// TIA Portal project "HR001_PLC_20260509" (V19)

(* hardware
DEVICE "S7-1200 station_1"  SIMATIC 1200-Station
   slot 0: "S7-1200 rack"  Rack  V1.0
   slot 1: "CPU_1200"  CPU 1215C DC/DC/DC  6ES7 215-1AG40-0XB0  V4.4
   slot 2: "DI 16/DQ 16x24VDC_1"  6ES7 223-1BL32-0XB0  V2.0
   slot 3: "DI 16/DQ 16x24VDC_2"  6ES7 223-1BL32-0XB0  V2.0
   slot 4: "DI 16x24VDC_1"  6ES7 221-1BH32-0XB0  V2.0
DEVICE "GSD device_11"  GSD.Device.PN
   slot 0: "机架"  Rack  V1.0
   slot 0: "AG1521Kuka_Big"  KRC4-ProfiNet_3.2  V3.2
      slot 0: "KRC4-ProfiNet_3.2"  KRC4-ProfiNet_3.2
      slot 1: "Interface1"  Interface1
         slot 1: "Port1"  Port1
   slot 2: "512 digital in- and outputs_1"  512 digital in- and outputs  KUKA KR C4 Device IO512
      slot 0: "512 digital in- and outputs"  512 digital in- and outputs
DEVICE "TP"  SIMATIC PC station
   slot 0: "HMI"  Rail  SIMATIC PC-Station  V1.0
      slot 125: "Stationmanager"  Station_Manager  V6.0.4
   slot 1: "HMI_RT_1"  WinCC RT Advanced  6AV2 104-0xxxx-xxxx  16.0.0.0
      slot 33792: "Computer interface"  Host interface
   slot 4: "IE general_1"  IE General  IE_CP  V8.2.0
*)

// ===== PLC "CPU_1200"  CPU 1215C DC/DC/DC =====
// protected blocks, not shown: "FB1003_CR", "FC1003_CR"

VAR_GLOBAL   // PLC tag table "M变量"
   "ManMode_M" AT %M26.0 : Bool;   // 手动模式
   "MastMode_M" AT %M26.1 : Bool;   // 校验模式
   "StepMode_M" AT %M26.2 : Bool;   // 单步模式
   "AutoMode_M" AT %M26.3 : Bool;   // 自动模式
   "EMMode_M" AT %M26.4 : Bool;   // 急停
   "StepPls_M" AT %M26.5 : Bool;   // 单步
   "AutoModeStarted_M" AT %M26.7 : Bool;   // 自动开始
   "ASMode_M" AT %M27.0 : Bool;   // 自动、单步
   "ASMMode_M" AT %M27.1 : Bool;   // 自动、单步、校验模式
   "AllMode_M" AT %M27.2 : Bool;   // 所有模式
   "ErrRst_M" AT %M27.3 : Bool;   // 故障复位
   "ErrRst_M_Auto" AT %M27.4 : Bool;   // 故障复位(系统参数可以设置为自动复位信号)
   "TRUE" AT %M29.0 : Bool;
   "False" AT %M29.1 : Bool;
   "MESConnect" AT %M29.3 : Bool;   // 0单机1联机
   "Debug_True" AT %M29.4 : Bool;   // 调试的时候，临时关闭
   "SyS_Time" AT %MD30 : Time_Of_Day;
   "Tag_1" AT %MW120 : Word;
   "Tag_2" AT %MW108 : Word;
   "Tag_3" AT %MW112 : UInt;
   "Tag_4" AT %M29.5 : Bool;
END_VAR

VAR_GLOBAL   // PLC tag table "PLC_IO"
   "IDoor3Unlocked" AT %I2.0 : Bool;   // 垂直击打门锁未锁定
   "IDoor3Insert" AT %I2.1 : Bool;   // 垂直击打门锁已插入
   "AStation_ToolOn2" AT %I2.5 : Bool;   // A工位夹具 有无检测2
   "AStation_ToolOn1" AT %I2.4 : Bool;   // A工位夹具 有无检测1
   "AStation_IZ03ExtPos" AT %I3.0 : Bool;   // A工位 旋转压紧缸伸出磁开
   "AStation_IZ03RetPos" AT %I3.1 : Bool;   // A工位 旋转压紧缸缩回磁开
   "BStation_ToolOn2" AT %I2.3 : Bool;   // B工位夹具有无检测2
   "BStation_ToolOn1" AT %I2.2 : Bool;   // B工位夹具 有无检测1
   "ICurtainErrRst" AT %I1.0 : Bool;   // 光幕复位按钮
   "IDoorOverRide" AT %I1.1 : Bool;   // 安全门旁路
   "IDoor1Unlocked" AT %I1.2 : Bool;   // 产品上料门锁未锁定
   "IDoor1Insert" AT %I1.3 : Bool;   // 产品上料门锁已插入
   "IDoor2Unlocked" AT %I1.4 : Bool;   // 水平击打门锁未锁定
   "IDoor2Insert" AT %I1.5 : Bool;   // 水平击打门锁已插入
   "IFixtureCode02" AT %I4.0 : Bool;   // 夹具电源快插编码2
   "IFixtureCode03" AT %I4.1 : Bool;   // 夹具电源快插编码3
   "IFixtureIOCode01" AT %I4.2 : Bool;   // 夹具IO快插编码1
   "IFixtureIOCode02" AT %I4.3 : Bool;   // 夹具IO快插编码2
   "IFixtureIOCode03" AT %I4.4 : Bool;   // 夹具IO快插编码3
   "IEMClamp" AT %I4.5 : Bool;   // 夹具侧急停按钮
   "IFixtureStuckSensor" AT %I4.6 : Bool;   // 夹具防卡信号
   "ISp4_7" AT %I4.7 : Bool;
   "IRobotEMOK" AT %I5.1 : Bool;   // 机器人急停按钮OK
   "ICurtainsOK" AT %I0.6 : Bool;   // 光幕OK信号
   "BStation_IZ04RetPos" AT %I2.6 : Bool;   // B工位 旋转压紧缸缩回磁开
   "IZ02RetPos" AT %I3.3 : Bool;   // 辅助气缸缩回磁开
   "IZ07ExtPos" AT %I3.5 : Bool;   // 机器人快换盘夹紧
   "IZ07RetPos" AT %I3.4 : Bool;   // 机器人快换盘松开
   "IToolAtPos" AT %I3.6 : Bool;   // 机器人快换盘在位
   "IFixtureCode01" AT %I3.7 : Bool;   // 夹具电源快插编码1
   "IEMOK" AT %I0.0 : Bool;   // 紧急停止OK
   "IAirPressOK" AT %I0.1 : Bool;   // 总气压检测OK
   "IMan" AT %I0.2 : Bool;   // 手动模式
   "IAuto" AT %I0.3 : Bool;   // 自动模式
   "IAutoModeStart" AT %I0.4 : Bool;   // 自动启动按钮
   "IErrRst" AT %I0.5 : Bool;   // 故障复位按钮
   "BStation_IZ04ExtPos" AT %I2.7 : Bool;   // B工位 旋转压紧缸伸出磁开
   "IZ02ExtPos" AT %I3.2 : Bool;   // 辅助气缸伸出磁开
   "IAllDoorClose" AT %I5.0 : Bool;   // 上电&所有 安全门关闭
   "IEMOK1" AT %I0.7 : Bool;   // 操作盒急停OK
   "ITempErr" AT %I5.2 : Bool;   // 温控器报警
   "IInsideEMOK" AT %I5.3 : Bool;   // 围栏内侧急停信号
   "IInsideEMOK1" AT %I5.4 : Bool;   // 水泥块击打框架急停信号
   "ISp055" AT %I5.5 : Bool;   // 备用
   "ISp056" AT %I5.6 : Bool;   // 备用
   "ISp057" AT %I5.7 : Bool;   // 备用
   "QBeeper" AT %Q0.2 : Bool;   // 蜂鸣器
   "QPanelG" AT %Q0.0 : Bool;   // 绿色运行指示灯
   "QPanelRed" AT %Q0.1 : Bool;   // 故障复位红灯
   "QTLR" AT %Q0.3 : Bool;   // 五色塔灯(红)
   "QTLY" AT %Q0.4 : Bool;   // 五色塔灯(黄)
   "QTLG" AT %Q0.5 : Bool;   // 五色塔灯(绿)
   "QTLB" AT %Q0.6 : Bool;   // 五色塔灯(蓝)
   "QTLW" AT %Q0.7 : Bool;   // 五色塔灯(白)
   "QSpairMode" AT %Q1.0 : Bool;   // 安全门旁路
   "QLampCtr" AT %Q1.1 : Bool;   // 日光灯控制中继（预留）
   "OOpenCamCover" AT %Q1.2 : Bool;   // 打开相机防护罩
   "OCloseCamCover" AT %Q1.3 : Bool;   // 关闭相机防护罩
   "QSp014" AT %Q1.4 : Bool;
   "QSp015" AT %Q1.5 : Bool;
   "QSp016" AT %Q1.6 : Bool;
   "QSp017" AT %Q1.7 : Bool;
   "QAStationFan" AT %Q3.5 : Bool;   // A Station Cooling Fan
   "QZ01RetEvt" AT %Q4.1 : Bool;   // Z1推力气缸缩回电磁阀
   "QZ02ExtEvt" AT %Q4.2 : Bool;   // Z2辅助气缸伸出电磁阀
   "QZ02RetEvt" AT %Q4.3 : Bool;   // Z2辅助气缸缩回电磁阀
   "QZ03ExtEvt" AT %Q4.4 : Bool;   // B工位防尘盖夹紧缸 伸出电磁阀
   "QZ03RetEvt" AT %Q4.5 : Bool;   // B工位左防尘盖夹紧缸 缩回电磁阀
   "QSpare026" AT %Q2.6 : Bool;
   "QCamCoverExt" AT %Q5.2 : Bool;   // 视觉保护罩气缸伸出
   "QSpare050" AT %Q5.0 : Bool;
   "DiamondVibCylinder" AT %Q5.1 : Bool;   // 水钻岩芯振动气缸
   "QSpare030" AT %Q3.2 : Bool;   // 备用
   "QBStationFan" AT %Q3.6 : Bool;   // B Station Cooling Fan
   "QWaterContactor" AT %Q3.4 : Bool;   // Water Drill Power Contactor
   "QWaterValve" AT %Q3.3 : Bool;   // Water Valve
   "QZ01ExtEvt" AT %Q4.0 : Bool;   // Z1推力气缸伸出电磁阀
   "QCamCoverRet" AT %Q5.3 : Bool;   // 视觉保护罩气缸缩回
   "QDoorClose" AT %Q2.0 : Bool;   // 门锁电源中继
   "QCurtainLight" AT %Q2.1 : Bool;   // 光幕复位指示灯
   "QCurtainRst" AT %Q2.2 : Bool;   // 光幕复位to安继
   "QSpare023" AT %Q2.3 : Bool;
   "QSpare025" AT %Q2.5 : Bool;
   "QSpare024" AT %Q2.4 : Bool;
   "QSpare027" AT %Q2.7 : Bool;
   "QSpare028" AT %Q3.0 : Bool;   // 备用
   "QSpare029" AT %Q3.1 : Bool;   // 备用
   "QZ04ExtEvt" AT %Q4.6 : Bool;   // A工位防尘盖夹紧缸 伸出电磁阀
   "QZ04RetEvt" AT %Q4.7 : Bool;   // A工位防尘盖夹紧缸 缩回电磁阀
   "QCStationFan" AT %Q3.7 : Bool;   // C Station Cooling Fan
   "QZ14ExtEvt" AT %Q5.4 : Bool;   // Z14三爪卡盘气缸伸出电磁阀
   "QZ14RetEvt" AT %Q5.5 : Bool;   // Z14三爪卡盘气缸缩回电磁阀
   "QZ07ExtEvt" AT %Q5.7 : Bool;   // Z7快换盘锁紧电磁阀
   "QZ07RetEvt" AT %Q5.6 : Bool;   // Z7快换盘松开电磁阀
   "ISp060" AT %I6.0 : Bool;
   "ISp061" AT %I6.1 : Bool;
   "ISp062" AT %I6.2 : Bool;
   "ISp063" AT %I6.3 : Bool;
   "ISp064" AT %I6.4 : Bool;
   "ISp065" AT %I6.5 : Bool;
   "IW10" AT %IW10 : Int;   // 比例阀输出
   "QW10" AT %QW10 : Int;
   "IW12" AT %IW12 : Int;   // 推力缸长度
   "ISp066" AT %I6.6 : Bool;
   "ISp067" AT %I6.7 : Bool;
   "ICoreBlockDect_LeftTool" AT %I7.0 : Bool;   // 左侧水钻工具岩心检测
   "ICoreBlockDect_RightTool" AT %I7.1 : Bool;   // 右侧水钻工具岩心检测
   "IWaterToolAtDectPos" AT %I7.2 : Bool;   // 水钻工具到达检测位
   "ICoreBlockDropDect_LeftTool" AT %I7.3 : Bool;   // 左侧水钻工具岩心掉落检测
   "ICoreBlockDropDect_RightTool" AT %I7.4 : Bool;   // 右侧水钻工具岩心掉落检测
   "ISp075" AT %I7.5 : Bool;
   "ISp076" AT %I7.6 : Bool;
   "ISp077" AT %I7.7 : Bool;
END_VAR

TYPE "UDT_Step"
VERSION : 0.1
   STRUCT
      StartCmd_ManMode : Bool;   // DoManual
      StartCmd_AutoMode : Bool;   // 自动运行启动命令；
      OkToStart : Bool;   // 条件满足，允许启动
      HomePos : Bool;   // 工位在原点位置
      "Do" : Bool;   // 本工位必须要做(可能条件暂时不满足)
      Done : Bool;   // 工位完成信号
      PartOn : Bool;   // 有工件标志
      PartOK : Bool;   // 产品合格标志
      PartNG : Bool;   // 产品不合格标志
      Start : Bool;
      End : Bool;
      ErrEnd : Bool;
      S1 : Bool;
      S2 : Bool;
      S3 : Bool;
      S4 : Bool;
      S5 : Bool;
      S6 : Bool;
      S7 : Bool;
      S8 : Bool;
      S9 : Bool;
      S10 : Bool;
      S11 : Bool;
      S12 : Bool;
      S13 : Bool;
      S14 : Bool;
      S15 : Bool;
      S16 : Bool;
      S17 : Bool;
      S18 : Bool;
      S19 : Bool;
      S20 : Bool;
      S21 : Bool;
      S22 : Bool;
      S23 : Bool;
      S24 : Bool;
      S25 : Bool;
      S26 : Bool;
      S27 : Bool;
      S28 : Bool;
      S29 : Bool;
      S30 : Bool;
      S31 : Bool;
      S32 : Bool;
      S33 : Bool;
      S34 : Bool;
      S35 : Bool;
      S36 : Bool;
      S37 : Bool;
      S38 : Bool;
      S39 : Bool;
      S40 : Bool;
      S41 : Bool;
      S42 : Bool;
      S43 : Bool;
      S44 : Bool;
      S45 : Bool;
      S46 : Bool;
      S47 : Bool;
      S48 : Bool;
      S49 : Bool;
      S50 : Bool;
      S51 : Bool;
      S52 : Bool;
      S53 : Bool;
      S54 : Bool;
      S55 : Bool;
      S56 : Bool;
      S57 : Bool;
      S58 : Bool;
      S59 : Bool;
      S60 : Bool;
      S61 : Bool;
      S62 : Bool;
      S63 : Bool;
      S64 : Bool;
      S65 : Bool;
      S66 : Bool;
      S67 : Bool;
   END_STRUCT;
END_TYPE

TYPE "UDT_DrillData"
   STRUCT
      CurrentDrillWidth : Real;   // 当前钻孔宽度 mm
      CurrentDrillLength : Real;   // 当前钻孔长度 mm
      CurrentDrillDepth : Real;   // 当前钻孔深度 mm
      LastDrillWidth : Real;   // 前钻孔宽度 mm
      LastDrillDepth : Real;   // 前钻孔深度 mm
      AlreadyDrillWidth : Real;   // 已钻宽度
      AlreadyDrillLength : Real;   // 已钻长度
      MaxWidth : Real;   // 当排最大钻孔宽度
      gi_OffsetX : Real;   // X方向偏移值
      gi_OffSetY : Real;   // Y方向偏移值
      gi_OffSetZ : Real;   // Z方向偏移值
      SlabWidth : Real;   // 水泥板宽度
      SlabLength : Real;   // 水泥板长度
      PosNo : Int;   // 孔位
      OppositeStartPos : Real;   // 反向开始坐标记忆
   END_STRUCT;
END_TYPE

// folder: 001_Para

TYPE "UDT_SystemPara"
VERSION : 0.1
   STRUCT
      bit : Struct
         ErrAutoResetOption : Bool;   // 故障自动复位功能
         MESActive : Bool;   // MES使能（1使能0屏蔽）
         sp : Word;
      END_STRUCT;
      Other : Struct
         OUT_Gain : Real;
         OUT_Offset : Real;
         IN_Gain : Real;
         IN_Offset : Real;
         IN_Gain_1 : Real;
         IN_Offset_1 : Real;
         sp : Array[0..191] of Byte;
      END_STRUCT;
   END_STRUCT;
END_TYPE

TYPE "UDT_TypePara"
VERSION : 0.1
   STRUCT
      TypeName : String[20];
      bit : Struct
         Bit0 : Bool;
         sp : Word;
         Other : Struct
            Bool_1 : Bool;   // ****功能选择（0：关闭，1：打开）
            Byte_2 : Byte;   // ****夹具编码（1~7）
            Int_1 : Int;   // ****读码长度（1~7）
            "Char" : Char;   // ****读码首字符
         END_STRUCT;
      END_STRUCT;
      Other : Struct
         STxxxCCDProgNO : Int;   // xxx功能相机程序号
         FixtureEnable : Bool;   // ****功能选择（0：关闭，1：打开）
         Byte_1 : Byte;   // ****夹具编码（1~7）
         Int_1 : Int;   // ****读码长度（1~7）
         "Char" : Char;   // ****读码首字符
         Word_1 : Word;   // ****夹具编码Word（1~7）
         DInt_1 : DInt;   // ****夹具编码DINT（1~7）
         DWord_1 : DWord;   // ****夹具编码DWord（1~7）
         Real_1 : Real;   // ****高度上限（1~7）
         S5Time : Time;   // ***延时（0.1~2.0）
         "String" : String[5];   // ***对比字符串
      END_STRUCT;
   END_STRUCT;
END_TYPE

// folder: (top level)

DATA_BLOCK "DB1001_SysMode"   // DB1001
{ S7_Optimized_Access := 'TRUE' }
VERSION : 0.1
// stored: InstanceOfName FB1001_SysMode
"FB1001_SysMode"
BEGIN
END_DATA_BLOCK

DATA_BLOCK "DB1010_Parameter"   // DB1010
{ S7_Optimized_Access := 'TRUE' }
VERSION : 0.1
// stored: InstanceOfName FB1010_Parameter
"FB1010_Parameter"
BEGIN
   SystemParaR.Other.OUT_Gain := 2.065072E-05;
   SystemParaR.Other.OUT_Offset := -0.00368739;
   SystemParaR.Other.IN_Gain := 757.8949;
   SystemParaR.Other.IN_Offset := -356.6613;
   SystemParaR.Other.IN_Gain_1 := -113.0993;
   SystemParaR.Other.IN_Offset_1 := 103.8807;
END_DATA_BLOCK

DATA_BLOCK "DB1089_AddrRegister"   // DB1089
{ S7_Optimized_Access := 'TRUE' }
VERSION : 0.1
// stored: InstanceOfName FB1089_AddrRegister
"FB1089_AddrRegister"
BEGIN
END_DATA_BLOCK

DATA_BLOCK "DB5000_ParameterLoadMemory"   // DB5000
{ S7_Optimized_Access := 'FALSE' }
VERSION : 0.1
   VAR
      SystemParaE : "UDT_SystemPara";
      AryTypePara : Array[0..300] of "UDT_TypePara";
      lastBit : Byte := 16#00;
   END_VAR
BEGIN
   AryTypePara[1].TypeName := '001';
   AryTypePara[1].Other.STxxxCCDProgNO := 1;
   AryTypePara[2].TypeName := '002';
   AryTypePara[2].Other.STxxxCCDProgNO := 2;
   AryTypePara[100].TypeName := '100';
   AryTypePara[100].Other.STxxxCCDProgNO := 100;
   AryTypePara[101].TypeName := '101';
   AryTypePara[101].Other.STxxxCCDProgNO := 101;
   AryTypePara[102].TypeName := '102';
   AryTypePara[102].Other.STxxxCCDProgNO := 102;
   AryTypePara[103].TypeName := '103';
   AryTypePara[103].Other.STxxxCCDProgNO := 103;
   AryTypePara[298].TypeName := '298';
   AryTypePara[298].Other.STxxxCCDProgNO := 300;
   AryTypePara[299].TypeName := '299';
   AryTypePara[299].Other.STxxxCCDProgNO := 299;
   AryTypePara[300].TypeName := '300';
   AryTypePara[300].Other.STxxxCCDProgNO := 300;
   AryTypePara[3].TypeName := '003';
   AryTypePara[4].TypeName := '004';
   AryTypePara[4].Other.STxxxCCDProgNO := 4;
   SystemParaE.bit.ErrAutoResetOption := FALSE;
   SystemParaE.bit.MESActive := FALSE;
   SystemParaE.bit.sp := 16#0000;
   SystemParaE.Other.OUT_Gain := 2.065072E-05;
   SystemParaE.Other.OUT_Offset := -0.00368739;
   SystemParaE.Other.IN_Gain := 757.8949;
   SystemParaE.Other.IN_Offset := -356.6613;
   SystemParaE.Other.IN_Gain_1 := -113.0993;
   SystemParaE.Other.IN_Offset_1 := 103.8807;
   SystemParaE.Other.sp[0] := 16#00;
   SystemParaE.Other.sp[1] := 16#00;
   SystemParaE.Other.sp[2] := 16#00;
   SystemParaE.Other.sp[3] := 16#00;
   SystemParaE.Other.sp[4] := 16#00;
   SystemParaE.Other.sp[5] := 16#00;
   SystemParaE.Other.sp[6] := 16#00;
   SystemParaE.Other.sp[7] := 16#00;
   SystemParaE.Other.sp[8] := 16#00;
   SystemParaE.Other.sp[9] := 16#00;
   SystemParaE.Other.sp[10] := 16#00;
   SystemParaE.Other.sp[11] := 16#00;
   SystemParaE.Other.sp[12] := 16#00;
   SystemParaE.Other.sp[13] := 16#00;
   SystemParaE.Other.sp[14] := 16#00;
   SystemParaE.Other.sp[15] := 16#00;
   SystemParaE.Other.sp[16] := 16#00;
   SystemParaE.Other.sp[17] := 16#00;
   SystemParaE.Other.sp[18] := 16#00;
   SystemParaE.Other.sp[19] := 16#00;
   SystemParaE.Other.sp[20] := 16#00;
   SystemParaE.Other.sp[21] := 16#00;
   SystemParaE.Other.sp[22] := 16#00;
   SystemParaE.Other.sp[23] := 16#00;
   SystemParaE.Other.sp[24] := 16#00;
   SystemParaE.Other.sp[25] := 16#00;
   SystemParaE.Other.sp[26] := 16#00;
   SystemParaE.Other.sp[27] := 16#00;
   SystemParaE.Other.sp[28] := 16#00;
   SystemParaE.Other.sp[29] := 16#00;
   SystemParaE.Other.sp[30] := 16#00;
   SystemParaE.Other.sp[31] := 16#00;
   SystemParaE.Other.sp[32] := 16#00;
   SystemParaE.Other.sp[33] := 16#00;
   SystemParaE.Other.sp[34] := 16#00;
   SystemParaE.Other.sp[35] := 16#00;
   SystemParaE.Other.sp[36] := 16#00;
   SystemParaE.Other.sp[37] := 16#00;
   SystemParaE.Other.sp[38] := 16#00;
   SystemParaE.Other.sp[39] := 16#00;
   SystemParaE.Other.sp[40] := 16#00;
   SystemParaE.Other.sp[41] := 16#00;
   SystemParaE.Other.sp[42] := 16#00;
   SystemParaE.Other.sp[43] := 16#00;
   SystemParaE.Other.sp[44] := 16#00;
   SystemParaE.Other.sp[45] := 16#00;
   SystemParaE.Other.sp[46] := 16#00;
   SystemParaE.Other.sp[47] := 16#00;
   SystemParaE.Other.sp[48] := 16#00;
   SystemParaE.Other.sp[49] := 16#00;
   SystemParaE.Other.sp[50] := 16#00;
   SystemParaE.Other.sp[51] := 16#00;
   SystemParaE.Other.sp[52] := 16#00;
   SystemParaE.Other.sp[53] := 16#00;
   SystemParaE.Other.sp[54] := 16#00;
   SystemParaE.Other.sp[55] := 16#00;
   SystemParaE.Other.sp[56] := 16#00;
   SystemParaE.Other.sp[57] := 16#00;
   SystemParaE.Other.sp[58] := 16#00;
   SystemParaE.Other.sp[59] := 16#00;
   SystemParaE.Other.sp[60] := 16#00;
   SystemParaE.Other.sp[61] := 16#00;
   SystemParaE.Other.sp[62] := 16#00;
   SystemParaE.Other.sp[63] := 16#00;
   SystemParaE.Other.sp[64] := 16#00;
   SystemParaE.Other.sp[65] := 16#00;
   SystemParaE.Other.sp[66] := 16#00;
   SystemParaE.Other.sp[67] := 16#00;
   SystemParaE.Other.sp[68] := 16#00;
   SystemParaE.Other.sp[69] := 16#00;
   SystemParaE.Other.sp[70] := 16#00;
   SystemParaE.Other.sp[71] := 16#00;
   SystemParaE.Other.sp[72] := 16#00;
   SystemParaE.Other.sp[73] := 16#00;
   SystemParaE.Other.sp[74] := 16#00;
   SystemParaE.Other.sp[75] := 16#00;
   SystemParaE.Other.sp[76] := 16#00;
   SystemParaE.Other.sp[77] := 16#00;
   SystemParaE.Other.sp[78] := 16#00;
   SystemParaE.Other.sp[79] := 16#00;
   SystemParaE.Other.sp[80] := 16#00;
   SystemParaE.Other.sp[81] := 16#00;
   SystemParaE.Other.sp[82] := 16#00;
   SystemParaE.Other.sp[83] := 16#00;
   SystemParaE.Other.sp[84] := 16#00;
   SystemParaE.Other.sp[85] := 16#00;
   SystemParaE.Other.sp[86] := 16#00;
   SystemParaE.Other.sp[87] := 16#00;
   SystemParaE.Other.sp[88] := 16#00;
   SystemParaE.Other.sp[89] := 16#00;
   SystemParaE.Other.sp[90] := 16#00;
   SystemParaE.Other.sp[91] := 16#00;
   SystemParaE.Other.sp[92] := 16#00;
   SystemParaE.Other.sp[93] := 16#00;
   SystemParaE.Other.sp[94] := 16#00;
   SystemParaE.Other.sp[95] := 16#00;
   SystemParaE.Other.sp[96] := 16#00;
   SystemParaE.Other.sp[97] := 16#00;
   SystemParaE.Other.sp[98] := 16#00;
   SystemParaE.Other.sp[99] := 16#00;
   SystemParaE.Other.sp[100] := 16#00;
   SystemParaE.Other.sp[101] := 16#00;
   SystemParaE.Other.sp[102] := 16#00;
   SystemParaE.Other.sp[103] := 16#00;
   SystemParaE.Other.sp[104] := 16#00;
   SystemParaE.Other.sp[105] := 16#00;
   SystemParaE.Other.sp[106] := 16#00;
   SystemParaE.Other.sp[107] := 16#00;
   SystemParaE.Other.sp[108] := 16#00;
   SystemParaE.Other.sp[109] := 16#00;
   SystemParaE.Other.sp[110] := 16#00;
   SystemParaE.Other.sp[111] := 16#00;
   SystemParaE.Other.sp[112] := 16#00;
   SystemParaE.Other.sp[113] := 16#00;
   SystemParaE.Other.sp[114] := 16#00;
   SystemParaE.Other.sp[115] := 16#00;
   SystemParaE.Other.sp[116] := 16#00;
   SystemParaE.Other.sp[117] := 16#00;
   SystemParaE.Other.sp[118] := 16#00;
   SystemParaE.Other.sp[119] := 16#00;
   SystemParaE.Other.sp[120] := 16#00;
   SystemParaE.Other.sp[121] := 16#00;
   SystemParaE.Other.sp[122] := 16#00;
   SystemParaE.Other.sp[123] := 16#00;
   SystemParaE.Other.sp[124] := 16#00;
   SystemParaE.Other.sp[125] := 16#00;
   SystemParaE.Other.sp[126] := 16#00;
   SystemParaE.Other.sp[127] := 16#00;
   SystemParaE.Other.sp[128] := 16#00;
   SystemParaE.Other.sp[129] := 16#00;
   SystemParaE.Other.sp[130] := 16#00;
   SystemParaE.Other.sp[131] := 16#00;
   SystemParaE.Other.sp[132] := 16#00;
   SystemParaE.Other.sp[133] := 16#00;
   SystemParaE.Other.sp[134] := 16#00;
   SystemParaE.Other.sp[135] := 16#00;
   SystemParaE.Other.sp[136] := 16#00;
   SystemParaE.Other.sp[137] := 16#00;
   SystemParaE.Other.sp[138] := 16#00;
   SystemParaE.Other.sp[139] := 16#00;
   SystemParaE.Other.sp[140] := 16#00;
   SystemParaE.Other.sp[141] := 16#00;
   SystemParaE.Other.sp[142] := 16#00;
   SystemParaE.Other.sp[143] := 16#00;
   SystemParaE.Other.sp[144] := 16#00;
   SystemParaE.Other.sp[145] := 16#00;
   SystemParaE.Other.sp[146] := 16#00;
   SystemParaE.Other.sp[147] := 16#00;
   SystemParaE.Other.sp[148] := 16#00;
   SystemParaE.Other.sp[149] := 16#00;
   SystemParaE.Other.sp[150] := 16#00;
   SystemParaE.Other.sp[151] := 16#00;
   SystemParaE.Other.sp[152] := 16#00;
   SystemParaE.Other.sp[153] := 16#00;
   SystemParaE.Other.sp[154] := 16#00;
   SystemParaE.Other.sp[155] := 16#00;
   SystemParaE.Other.sp[156] := 16#00;
   SystemParaE.Other.sp[157] := 16#00;
   SystemParaE.Other.sp[158] := 16#00;
   SystemParaE.Other.sp[159] := 16#00;
   SystemParaE.Other.sp[160] := 16#00;
   SystemParaE.Other.sp[161] := 16#00;
   SystemParaE.Other.sp[162] := 16#00;
   SystemParaE.Other.sp[163] := 16#00;
   SystemParaE.Other.sp[164] := 16#00;
   SystemParaE.Other.sp[165] := 16#00;
   SystemParaE.Other.sp[166] := 16#00;
   SystemParaE.Other.sp[167] := 16#00;
   SystemParaE.Other.sp[168] := 16#00;
   SystemParaE.Other.sp[169] := 16#00;
   SystemParaE.Other.sp[170] := 16#00;
   SystemParaE.Other.sp[171] := 16#00;
   SystemParaE.Other.sp[172] := 16#00;
   SystemParaE.Other.sp[173] := 16#00;
   SystemParaE.Other.sp[174] := 16#00;
   SystemParaE.Other.sp[175] := 16#00;
   SystemParaE.Other.sp[176] := 16#00;
   SystemParaE.Other.sp[177] := 16#00;
   SystemParaE.Other.sp[178] := 16#00;
   SystemParaE.Other.sp[179] := 16#00;
   SystemParaE.Other.sp[180] := 16#00;
   SystemParaE.Other.sp[181] := 16#00;
   SystemParaE.Other.sp[182] := 16#00;
   SystemParaE.Other.sp[183] := 16#00;
   SystemParaE.Other.sp[184] := 16#00;
   SystemParaE.Other.sp[185] := 16#00;
   SystemParaE.Other.sp[186] := 16#00;
   SystemParaE.Other.sp[187] := 16#00;
   SystemParaE.Other.sp[188] := 16#00;
   SystemParaE.Other.sp[189] := 16#00;
   SystemParaE.Other.sp[190] := 16#00;
   SystemParaE.Other.sp[191] := 16#00;
   AryTypePara[0].TypeName := '';
   AryTypePara[0].bit.Bit0 := FALSE;
   AryTypePara[0].bit.sp := 16#0000;
   AryTypePara[0].bit.Other.Bool_1 := FALSE;
   AryTypePara[0].bit.Other.Byte_2 := 16#00;
   AryTypePara[0].bit.Other.Int_1 := 0;
   AryTypePara[0].bit.Other."Char" := ' ';
   AryTypePara[0].Other.STxxxCCDProgNO := 0;
   AryTypePara[0].Other.FixtureEnable := FALSE;
   AryTypePara[0].Other.Byte_1 := 16#00;
   AryTypePara[0].Other.Int_1 := 0;
   AryTypePara[0].Other."Char" := ' ';
   AryTypePara[0].Other.Word_1 := 16#0000;
   AryTypePara[0].Other.DInt_1 := 0;
   AryTypePara[0].Other.DWord_1 := 16#0000_0000;
   AryTypePara[0].Other.Real_1 := 0.0;
   AryTypePara[0].Other.S5Time := T#0MS;
   AryTypePara[0].Other."String" := '';
   AryTypePara[1].bit.Bit0 := FALSE;
   AryTypePara[1].bit.sp := 16#0000;
   AryTypePara[1].bit.Other.Bool_1 := FALSE;
   AryTypePara[1].bit.Other.Byte_2 := 16#00;
   AryTypePara[1].bit.Other.Int_1 := 0;
   AryTypePara[1].bit.Other."Char" := ' ';
   AryTypePara[1].Other.FixtureEnable := FALSE;
   AryTypePara[1].Other.Byte_1 := 16#00;
   AryTypePara[1].Other.Int_1 := 0;
   AryTypePara[1].Other."Char" := ' ';
   AryTypePara[1].Other.Word_1 := 16#0000;
   AryTypePara[1].Other.DInt_1 := 0;
   AryTypePara[1].Other.DWord_1 := 16#0000_0000;
   AryTypePara[1].Other.Real_1 := 0.0;
   AryTypePara[1].Other.S5Time := T#0MS;
   AryTypePara[1].Other."String" := '';
   AryTypePara[2].bit.Bit0 := FALSE;
   AryTypePara[2].bit.sp := 16#0000;
   AryTypePara[2].bit.Other.Bool_1 := FALSE;
   AryTypePara[2].bit.Other.Byte_2 := 16#00;
   AryTypePara[2].bit.Other.Int_1 := 0;
   AryTypePara[2].bit.Other."Char" := ' ';
   AryTypePara[2].Other.FixtureEnable := FALSE;
   AryTypePara[2].Other.Byte_1 := 16#00;
   AryTypePara[2].Other.Int_1 := 0;
   AryTypePara[2].Other."Char" := ' ';
   AryTypePara[2].Other.Word_1 := 16#0000;
   AryTypePara[2].Other.DInt_1 := 0;
   AryTypePara[2].Other.DWord_1 := 16#0000_0000;
   AryTypePara[2].Other.Real_1 := 0.0;
   AryTypePara[2].Other.S5Time := T#0MS;
   AryTypePara[2].Other."String" := '';
   AryTypePara[3].bit.Bit0 := FALSE;
   AryTypePara[3].bit.sp := 16#0000;
   AryTypePara[3].bit.Other.Bool_1 := FALSE;
   AryTypePara[3].bit.Other.Byte_2 := 16#00;
   AryTypePara[3].bit.Other.Int_1 := 0;
   AryTypePara[3].bit.Other."Char" := ' ';
   AryTypePara[3].Other.STxxxCCDProgNO := 0;
   AryTypePara[3].Other.FixtureEnable := FALSE;
   AryTypePara[3].Other.Byte_1 := 16#00;
   AryTypePara[3].Other.Int_1 := 0;
   AryTypePara[3].Other."Char" := ' ';
   AryTypePara[3].Other.Word_1 := 16#0000;
   AryTypePara[3].Other.DInt_1 := 0;
   AryTypePara[3].Other.DWord_1 := 16#0000_0000;
   AryTypePara[3].Other.Real_1 := 0.0;
   AryTypePara[3].Other.S5Time := T#0MS;
   AryTypePara[3].Other."String" := '';
   AryTypePara[4].bit.Bit0 := FALSE;
   AryTypePara[4].bit.sp := 16#0000;
   AryTypePara[4].bit.Other.Bool_1 := FALSE;
   AryTypePara[4].bit.Other.Byte_2 := 16#00;
   AryTypePara[4].bit.Other.Int_1 := 0;
   AryTypePara[4].bit.Other."Char" := ' ';
   AryTypePara[4].Other.FixtureEnable := FALSE;
   AryTypePara[4].Other.Byte_1 := 16#00;
   AryTypePara[4].Other.Int_1 := 0;
   AryTypePara[4].Other."Char" := ' ';
   AryTypePara[4].Other.Word_1 := 16#0000;
   AryTypePara[4].Other.DInt_1 := 0;
   AryTypePara[4].Other.DWord_1 := 16#0000_0000;
   AryTypePara[4].Other.Real_1 := 0.0;
   AryTypePara[4].Other.S5Time := T#0MS;
   AryTypePara[4].Other."String" := '';
   AryTypePara[5].TypeName := '';
   AryTypePara[5].bit.Bit0 := FALSE;
   AryTypePara[5].bit.sp := 16#0000;
   AryTypePara[5].bit.Other.Bool_1 := FALSE;
   AryTypePara[5].bit.Other.Byte_2 := 16#00;
   AryTypePara[5].bit.Other.Int_1 := 0;
   AryTypePara[5].bit.Other."Char" := ' ';
   AryTypePara[5].Other.STxxxCCDProgNO := 0;
   AryTypePara[5].Other.FixtureEnable := FALSE;
   AryTypePara[5].Other.Byte_1 := 16#00;
   AryTypePara[5].Other.Int_1 := 0;
   AryTypePara[5].Other."Char" := ' ';
   AryTypePara[5].Other.Word_1 := 16#0000;
   AryTypePara[5].Other.DInt_1 := 0;
   AryTypePara[5].Other.DWord_1 := 16#0000_0000;
   AryTypePara[5].Other.Real_1 := 0.0;
   AryTypePara[5].Other.S5Time := T#0MS;
   AryTypePara[5].Other."String" := '';
   AryTypePara[6].TypeName := '';
   AryTypePara[6].bit.Bit0 := FALSE;
   AryTypePara[6].bit.sp := 16#0000;
   AryTypePara[6].bit.Other.Bool_1 := FALSE;
   AryTypePara[6].bit.Other.Byte_2 := 16#00;
   AryTypePara[6].bit.Other.Int_1 := 0;
   AryTypePara[6].bit.Other."Char" := ' ';
   AryTypePara[6].Other.STxxxCCDProgNO := 0;
   AryTypePara[6].Other.FixtureEnable := FALSE;
   AryTypePara[6].Other.Byte_1 := 16#00;
   AryTypePara[6].Other.Int_1 := 0;
   AryTypePara[6].Other."Char" := ' ';
   AryTypePara[6].Other.Word_1 := 16#0000;
   AryTypePara[6].Other.DInt_1 := 0;
   AryTypePara[6].Other.DWord_1 := 16#0000_0000;
   AryTypePara[6].Other.Real_1 := 0.0;
   AryTypePara[6].Other.S5Time := T#0MS;
   AryTypePara[6].Other."String" := '';
   AryTypePara[7].TypeName := '';
   AryTypePara[7].bit.Bit0 := FALSE;
   AryTypePara[7].bit.sp := 16#0000;
   AryTypePara[7].bit.Other.Bool_1 := FALSE;
   AryTypePara[7].bit.Other.Byte_2 := 16#00;
   AryTypePara[7].bit.Other.Int_1 := 0;
   AryTypePara[7].bit.Other."Char" := ' ';
   AryTypePara[7].Other.STxxxCCDProgNO := 0;
   AryTypePara[7].Other.FixtureEnable := FALSE;
   AryTypePara[7].Other.Byte_1 := 16#00;
   AryTypePara[7].Other.Int_1 := 0;
   AryTypePara[7].Other."Char" := ' ';
   AryTypePara[7].Other.Word_1 := 16#0000;
   AryTypePara[7].Other.DInt_1 := 0;
   AryTypePara[7].Other.DWord_1 := 16#0000_0000;
   AryTypePara[7].Other.Real_1 := 0.0;
   AryTypePara[7].Other.S5Time := T#0MS;
   AryTypePara[7].Other."String" := '';
   AryTypePara[8].TypeName := '';
   AryTypePara[8].bit.Bit0 := FALSE;
   AryTypePara[8].bit.sp := 16#0000;
   AryTypePara[8].bit.Other.Bool_1 := FALSE;
   AryTypePara[8].bit.Other.Byte_2 := 16#00;
   AryTypePara[8].bit.Other.Int_1 := 0;
   AryTypePara[8].bit.Other."Char" := ' ';
   AryTypePara[8].Other.STxxxCCDProgNO := 0;
   AryTypePara[8].Other.FixtureEnable := FALSE;
   AryTypePara[8].Other.Byte_1 := 16#00;
   AryTypePara[8].Other.Int_1 := 0;
   AryTypePara[8].Other."Char" := ' ';
   AryTypePara[8].Other.Word_1 := 16#0000;
   AryTypePara[8].Other.DInt_1 := 0;
   AryTypePara[8].Other.DWord_1 := 16#0000_0000;
   AryTypePara[8].Other.Real_1 := 0.0;
   AryTypePara[8].Other.S5Time := T#0MS;
   AryTypePara[8].Other."String" := '';
   AryTypePara[9].TypeName := '';
   AryTypePara[9].bit.Bit0 := FALSE;
   AryTypePara[9].bit.sp := 16#0000;
   AryTypePara[9].bit.Other.Bool_1 := FALSE;
   AryTypePara[9].bit.Other.Byte_2 := 16#00;
   AryTypePara[9].bit.Other.Int_1 := 0;
   AryTypePara[9].bit.Other."Char" := ' ';
   AryTypePara[9].Other.STxxxCCDProgNO := 0;
   AryTypePara[9].Other.FixtureEnable := FALSE;
   AryTypePara[9].Other.Byte_1 := 16#00;
   AryTypePara[9].Other.Int_1 := 0;
   AryTypePara[9].Other."Char" := ' ';
   AryTypePara[9].Other.Word_1 := 16#0000;
   AryTypePara[9].Other.DInt_1 := 0;
   AryTypePara[9].Other.DWord_1 := 16#0000_0000;
   AryTypePara[9].Other.Real_1 := 0.0;
   AryTypePara[9].Other.S5Time := T#0MS;
   AryTypePara[9].Other."String" := '';
   AryTypePara[10].TypeName := '';
   AryTypePara[10].bit.Bit0 := FALSE;
   AryTypePara[10].bit.sp := 16#0000;
   AryTypePara[10].bit.Other.Bool_1 := FALSE;
   AryTypePara[10].bit.Other.Byte_2 := 16#00;
   AryTypePara[10].bit.Other.Int_1 := 0;
   AryTypePara[10].bit.Other."Char" := ' ';
   AryTypePara[10].Other.STxxxCCDProgNO := 0;
   AryTypePara[10].Other.FixtureEnable := FALSE;
   AryTypePara[10].Other.Byte_1 := 16#00;
   AryTypePara[10].Other.Int_1 := 0;
   AryTypePara[10].Other."Char" := ' ';
   AryTypePara[10].Other.Word_1 := 16#0000;
   AryTypePara[10].Other.DInt_1 := 0;
   AryTypePara[10].Other.DWord_1 := 16#0000_0000;
   AryTypePara[10].Other.Real_1 := 0.0;
   AryTypePara[10].Other.S5Time := T#0MS;
   AryTypePara[10].Other."String" := '';
   AryTypePara[11].TypeName := '';
   AryTypePara[11].bit.Bit0 := FALSE;
   AryTypePara[11].bit.sp := 16#0000;
   AryTypePara[11].bit.Other.Bool_1 := FALSE;
   AryTypePara[11].bit.Other.Byte_2 := 16#00;
   AryTypePara[11].bit.Other.Int_1 := 0;
   AryTypePara[11].bit.Other."Char" := ' ';
   AryTypePara[11].Other.STxxxCCDProgNO := 0;
   AryTypePara[11].Other.FixtureEnable := FALSE;
   AryTypePara[11].Other.Byte_1 := 16#00;
   AryTypePara[11].Other.Int_1 := 0;
   AryTypePara[11].Other."Char" := ' ';
   AryTypePara[11].Other.Word_1 := 16#0000;
   AryTypePara[11].Other.DInt_1 := 0;
   AryTypePara[11].Other.DWord_1 := 16#0000_0000;
   AryTypePara[11].Other.Real_1 := 0.0;
   AryTypePara[11].Other.S5Time := T#0MS;
   AryTypePara[11].Other."String" := '';
   AryTypePara[12].TypeName := '';
   AryTypePara[12].bit.Bit0 := FALSE;
   AryTypePara[12].bit.sp := 16#0000;
   AryTypePara[12].bit.Other.Bool_1 := FALSE;
   AryTypePara[12].bit.Other.Byte_2 := 16#00;
   AryTypePara[12].bit.Other.Int_1 := 0;
   AryTypePara[12].bit.Other."Char" := ' ';
   AryTypePara[12].Other.STxxxCCDProgNO := 0;
   AryTypePara[12].Other.FixtureEnable := FALSE;
   AryTypePara[12].Other.Byte_1 := 16#00;
   AryTypePara[12].Other.Int_1 := 0;
   AryTypePara[12].Other."Char" := ' ';
   AryTypePara[12].Other.Word_1 := 16#0000;
   AryTypePara[12].Other.DInt_1 := 0;
   AryTypePara[12].Other.DWord_1 := 16#0000_0000;
   AryTypePara[12].Other.Real_1 := 0.0;
   AryTypePara[12].Other.S5Time := T#0MS;
   AryTypePara[12].Other."String" := '';
   AryTypePara[13].TypeName := '';
   AryTypePara[13].bit.Bit0 := FALSE;
   AryTypePara[13].bit.sp := 16#0000;
   AryTypePara[13].bit.Other.Bool_1 := FALSE;
   AryTypePara[13].bit.Other.Byte_2 := 16#00;
   AryTypePara[13].bit.Other.Int_1 := 0;
   AryTypePara[13].bit.Other."Char" := ' ';
   AryTypePara[13].Other.STxxxCCDProgNO := 0;
   AryTypePara[13].Other.FixtureEnable := FALSE;
   AryTypePara[13].Other.Byte_1 := 16#00;
   AryTypePara[13].Other.Int_1 := 0;
   AryTypePara[13].Other."Char" := ' ';
   AryTypePara[13].Other.Word_1 := 16#0000;
   AryTypePara[13].Other.DInt_1 := 0;
   AryTypePara[13].Other.DWord_1 := 16#0000_0000;
   AryTypePara[13].Other.Real_1 := 0.0;
   AryTypePara[13].Other.S5Time := T#0MS;
   AryTypePara[13].Other."String" := '';
   AryTypePara[14].TypeName := '';
   AryTypePara[14].bit.Bit0 := FALSE;
   AryTypePara[14].bit.sp := 16#0000;
   AryTypePara[14].bit.Other.Bool_1 := FALSE;
   AryTypePara[14].bit.Other.Byte_2 := 16#00;
   AryTypePara[14].bit.Other.Int_1 := 0;
   AryTypePara[14].bit.Other."Char" := ' ';
   AryTypePara[14].Other.STxxxCCDProgNO := 0;
   AryTypePara[14].Other.FixtureEnable := FALSE;
   AryTypePara[14].Other.Byte_1 := 16#00;
   AryTypePara[14].Other.Int_1 := 0;
   AryTypePara[14].Other."Char" := ' ';
   AryTypePara[14].Other.Word_1 := 16#0000;
   AryTypePara[14].Other.DInt_1 := 0;
   AryTypePara[14].Other.DWord_1 := 16#0000_0000;
   AryTypePara[14].Other.Real_1 := 0.0;
   AryTypePara[14].Other.S5Time := T#0MS;
   AryTypePara[14].Other."String" := '';
   AryTypePara[15].TypeName := '';
   AryTypePara[15].bit.Bit0 := FALSE;
   AryTypePara[15].bit.sp := 16#0000;
   AryTypePara[15].bit.Other.Bool_1 := FALSE;
   AryTypePara[15].bit.Other.Byte_2 := 16#00;
   AryTypePara[15].bit.Other.Int_1 := 0;
   AryTypePara[15].bit.Other."Char" := ' ';
   AryTypePara[15].Other.STxxxCCDProgNO := 0;
   AryTypePara[15].Other.FixtureEnable := FALSE;
   AryTypePara[15].Other.Byte_1 := 16#00;
   AryTypePara[15].Other.Int_1 := 0;
   AryTypePara[15].Other."Char" := ' ';
   AryTypePara[15].Other.Word_1 := 16#0000;
   AryTypePara[15].Other.DInt_1 := 0;
   AryTypePara[15].Other.DWord_1 := 16#0000_0000;
   AryTypePara[15].Other.Real_1 := 0.0;
   AryTypePara[15].Other.S5Time := T#0MS;
   AryTypePara[15].Other."String" := '';
   AryTypePara[16].TypeName := '';
   AryTypePara[16].bit.Bit0 := FALSE;
   AryTypePara[16].bit.sp := 16#0000;
   AryTypePara[16].bit.Other.Bool_1 := FALSE;
   AryTypePara[16].bit.Other.Byte_2 := 16#00;
   AryTypePara[16].bit.Other.Int_1 := 0;
   AryTypePara[16].bit.Other."Char" := ' ';
   AryTypePara[16].Other.STxxxCCDProgNO := 0;
   AryTypePara[16].Other.FixtureEnable := FALSE;
   AryTypePara[16].Other.Byte_1 := 16#00;
   AryTypePara[16].Other.Int_1 := 0;
   AryTypePara[16].Other."Char" := ' ';
   AryTypePara[16].Other.Word_1 := 16#0000;
   AryTypePara[16].Other.DInt_1 := 0;
   AryTypePara[16].Other.DWord_1 := 16#0000_0000;
   AryTypePara[16].Other.Real_1 := 0.0;
   AryTypePara[16].Other.S5Time := T#0MS;
   AryTypePara[16].Other."String" := '';
   AryTypePara[17].TypeName := '';
   AryTypePara[17].bit.Bit0 := FALSE;
   AryTypePara[17].bit.sp := 16#0000;
   AryTypePara[17].bit.Other.Bool_1 := FALSE;
   AryTypePara[17].bit.Other.Byte_2 := 16#00;
   AryTypePara[17].bit.Other.Int_1 := 0;
   AryTypePara[17].bit.Other."Char" := ' ';
   AryTypePara[17].Other.STxxxCCDProgNO := 0;
   AryTypePara[17].Other.FixtureEnable := FALSE;
   AryTypePara[17].Other.Byte_1 := 16#00;
   AryTypePara[17].Other.Int_1 := 0;
   AryTypePara[17].Other."Char" := ' ';
   AryTypePara[17].Other.Word_1 := 16#0000;
   AryTypePara[17].Other.DInt_1 := 0;
   AryTypePara[17].Other.DWord_1 := 16#0000_0000;
   AryTypePara[17].Other.Real_1 := 0.0;
   AryTypePara[17].Other.S5Time := T#0MS;
   AryTypePara[17].Other."String" := '';
   AryTypePara[18].TypeName := '';
   AryTypePara[18].bit.Bit0 := FALSE;
   AryTypePara[18].bit.sp := 16#0000;
   AryTypePara[18].bit.Other.Bool_1 := FALSE;
   AryTypePara[18].bit.Other.Byte_2 := 16#00;
   AryTypePara[18].bit.Other.Int_1 := 0;
   AryTypePara[18].bit.Other."Char" := ' ';
   AryTypePara[18].Other.STxxxCCDProgNO := 0;
   AryTypePara[18].Other.FixtureEnable := FALSE;
   AryTypePara[18].Other.Byte_1 := 16#00;
   AryTypePara[18].Other.Int_1 := 0;
   AryTypePara[18].Other."Char" := ' ';
   AryTypePara[18].Other.Word_1 := 16#0000;
   AryTypePara[18].Other.DInt_1 := 0;
   AryTypePara[18].Other.DWord_1 := 16#0000_0000;
   AryTypePara[18].Other.Real_1 := 0.0;
   AryTypePara[18].Other.S5Time := T#0MS;
   AryTypePara[18].Other."String" := '';
   AryTypePara[19].TypeName := '';
   AryTypePara[19].bit.Bit0 := FALSE;
   AryTypePara[19].bit.sp := 16#0000;
   AryTypePara[19].bit.Other.Bool_1 := FALSE;
   AryTypePara[19].bit.Other.Byte_2 := 16#00;
   AryTypePara[19].bit.Other.Int_1 := 0;
   AryTypePara[19].bit.Other."Char" := ' ';
   AryTypePara[19].Other.STxxxCCDProgNO := 0;
   AryTypePara[19].Other.FixtureEnable := FALSE;
   AryTypePara[19].Other.Byte_1 := 16#00;
   AryTypePara[19].Other.Int_1 := 0;
   AryTypePara[19].Other."Char" := ' ';
   AryTypePara[19].Other.Word_1 := 16#0000;
   AryTypePara[19].Other.DInt_1 := 0;
   AryTypePara[19].Other.DWord_1 := 16#0000_0000;
   AryTypePara[19].Other.Real_1 := 0.0;
   AryTypePara[19].Other.S5Time := T#0MS;
   AryTypePara[19].Other."String" := '';
   AryTypePara[20].TypeName := '';
   AryTypePara[20].bit.Bit0 := FALSE;
   AryTypePara[20].bit.sp := 16#0000;
   AryTypePara[20].bit.Other.Bool_1 := FALSE;
   AryTypePara[20].bit.Other.Byte_2 := 16#00;
   AryTypePara[20].bit.Other.Int_1 := 0;
   AryTypePara[20].bit.Other."Char" := ' ';
   AryTypePara[20].Other.STxxxCCDProgNO := 0;
   AryTypePara[20].Other.FixtureEnable := FALSE;
   AryTypePara[20].Other.Byte_1 := 16#00;
   AryTypePara[20].Other.Int_1 := 0;
   AryTypePara[20].Other."Char" := ' ';
   AryTypePara[20].Other.Word_1 := 16#0000;
   AryTypePara[20].Other.DInt_1 := 0;
   AryTypePara[20].Other.DWord_1 := 16#0000_0000;
   AryTypePara[20].Other.Real_1 := 0.0;
   AryTypePara[20].Other.S5Time := T#0MS;
   AryTypePara[20].Other."String" := '';
   AryTypePara[21].TypeName := '';
   AryTypePara[21].bit.Bit0 := FALSE;
   AryTypePara[21].bit.sp := 16#0000;
   AryTypePara[21].bit.Other.Bool_1 := FALSE;
   AryTypePara[21].bit.Other.Byte_2 := 16#00;
   AryTypePara[21].bit.Other.Int_1 := 0;
   AryTypePara[21].bit.Other."Char" := ' ';
   AryTypePara[21].Other.STxxxCCDProgNO := 0;
   AryTypePara[21].Other.FixtureEnable := FALSE;
   AryTypePara[21].Other.Byte_1 := 16#00;
   AryTypePara[21].Other.Int_1 := 0;
   AryTypePara[21].Other."Char" := ' ';
   AryTypePara[21].Other.Word_1 := 16#0000;
   AryTypePara[21].Other.DInt_1 := 0;
   AryTypePara[21].Other.DWord_1 := 16#0000_0000;
   AryTypePara[21].Other.Real_1 := 0.0;
   AryTypePara[21].Other.S5Time := T#0MS;
   AryTypePara[21].Other."String" := '';
   AryTypePara[22].TypeName := '';
   AryTypePara[22].bit.Bit0 := FALSE;
   AryTypePara[22].bit.sp := 16#0000;
   AryTypePara[22].bit.Other.Bool_1 := FALSE;
   AryTypePara[22].bit.Other.Byte_2 := 16#00;
   AryTypePara[22].bit.Other.Int_1 := 0;
   AryTypePara[22].bit.Other."Char" := ' ';
   AryTypePara[22].Other.STxxxCCDProgNO := 0;
   AryTypePara[22].Other.FixtureEnable := FALSE;
   AryTypePara[22].Other.Byte_1 := 16#00;
   AryTypePara[22].Other.Int_1 := 0;
   AryTypePara[22].Other."Char" := ' ';
   AryTypePara[22].Other.Word_1 := 16#0000;
   AryTypePara[22].Other.DInt_1 := 0;
   AryTypePara[22].Other.DWord_1 := 16#0000_0000;
   AryTypePara[22].Other.Real_1 := 0.0;
   AryTypePara[22].Other.S5Time := T#0MS;
   AryTypePara[22].Other."String" := '';
   AryTypePara[23].TypeName := '';
   AryTypePara[23].bit.Bit0 := FALSE;
   AryTypePara[23].bit.sp := 16#0000;
   AryTypePara[23].bit.Other.Bool_1 := FALSE;
   AryTypePara[23].bit.Other.Byte_2 := 16#00;
   AryTypePara[23].bit.Other.Int_1 := 0;
   AryTypePara[23].bit.Other."Char" := ' ';
   AryTypePara[23].Other.STxxxCCDProgNO := 0;
   AryTypePara[23].Other.FixtureEnable := FALSE;
   AryTypePara[23].Other.Byte_1 := 16#00;
   AryTypePara[23].Other.Int_1 := 0;
   AryTypePara[23].Other."Char" := ' ';
   AryTypePara[23].Other.Word_1 := 16#0000;
   AryTypePara[23].Other.DInt_1 := 0;
   AryTypePara[23].Other.DWord_1 := 16#0000_0000;
   AryTypePara[23].Other.Real_1 := 0.0;
   AryTypePara[23].Other.S5Time := T#0MS;
   AryTypePara[23].Other."String" := '';
   AryTypePara[24].TypeName := '';
   AryTypePara[24].bit.Bit0 := FALSE;
   AryTypePara[24].bit.sp := 16#0000;
   AryTypePara[24].bit.Other.Bool_1 := FALSE;
   AryTypePara[24].bit.Other.Byte_2 := 16#00;
   AryTypePara[24].bit.Other.Int_1 := 0;
   AryTypePara[24].bit.Other."Char" := ' ';
   AryTypePara[24].Other.STxxxCCDProgNO := 0;
   AryTypePara[24].Other.FixtureEnable := FALSE;
   AryTypePara[24].Other.Byte_1 := 16#00;
   AryTypePara[24].Other.Int_1 := 0;
   AryTypePara[24].Other."Char" := ' ';
   AryTypePara[24].Other.Word_1 := 16#0000;
   AryTypePara[24].Other.DInt_1 := 0;
   AryTypePara[24].Other.DWord_1 := 16#0000_0000;
   AryTypePara[24].Other.Real_1 := 0.0;
   AryTypePara[24].Other.S5Time := T#0MS;
   AryTypePara[24].Other."String" := '';
   AryTypePara[25].TypeName := '';
   AryTypePara[25].bit.Bit0 := FALSE;
   AryTypePara[25].bit.sp := 16#0000;
   AryTypePara[25].bit.Other.Bool_1 := FALSE;
   AryTypePara[25].bit.Other.Byte_2 := 16#00;
   AryTypePara[25].bit.Other.Int_1 := 0;
   AryTypePara[25].bit.Other."Char" := ' ';
   AryTypePara[25].Other.STxxxCCDProgNO := 0;
   AryTypePara[25].Other.FixtureEnable := FALSE;
   AryTypePara[25].Other.Byte_1 := 16#00;
   AryTypePara[25].Other.Int_1 := 0;
   AryTypePara[25].Other."Char" := ' ';
   AryTypePara[25].Other.Word_1 := 16#0000;
   AryTypePara[25].Other.DInt_1 := 0;
   AryTypePara[25].Other.DWord_1 := 16#0000_0000;
   AryTypePara[25].Other.Real_1 := 0.0;
   AryTypePara[25].Other.S5Time := T#0MS;
   AryTypePara[25].Other."String" := '';
   AryTypePara[26].TypeName := '';
   AryTypePara[26].bit.Bit0 := FALSE;
   AryTypePara[26].bit.sp := 16#0000;
   AryTypePara[26].bit.Other.Bool_1 := FALSE;
   AryTypePara[26].bit.Other.Byte_2 := 16#00;
   AryTypePara[26].bit.Other.Int_1 := 0;
   AryTypePara[26].bit.Other."Char" := ' ';
   AryTypePara[26].Other.STxxxCCDProgNO := 0;
   AryTypePara[26].Other.FixtureEnable := FALSE;
   AryTypePara[26].Other.Byte_1 := 16#00;
   AryTypePara[26].Other.Int_1 := 0;
   AryTypePara[26].Other."Char" := ' ';
   AryTypePara[26].Other.Word_1 := 16#0000;
   AryTypePara[26].Other.DInt_1 := 0;
   AryTypePara[26].Other.DWord_1 := 16#0000_0000;
   AryTypePara[26].Other.Real_1 := 0.0;
   AryTypePara[26].Other.S5Time := T#0MS;
   AryTypePara[26].Other."String" := '';
   AryTypePara[27].TypeName := '';
   AryTypePara[27].bit.Bit0 := FALSE;
   AryTypePara[27].bit.sp := 16#0000;
   AryTypePara[27].bit.Other.Bool_1 := FALSE;
   AryTypePara[27].bit.Other.Byte_2 := 16#00;
   AryTypePara[27].bit.Other.Int_1 := 0;
   AryTypePara[27].bit.Other."Char" := ' ';
   AryTypePara[27].Other.STxxxCCDProgNO := 0;
   AryTypePara[27].Other.FixtureEnable := FALSE;
   AryTypePara[27].Other.Byte_1 := 16#00;
   AryTypePara[27].Other.Int_1 := 0;
   AryTypePara[27].Other."Char" := ' ';
   AryTypePara[27].Other.Word_1 := 16#0000;
   AryTypePara[27].Other.DInt_1 := 0;
   AryTypePara[27].Other.DWord_1 := 16#0000_0000;
   AryTypePara[27].Other.Real_1 := 0.0;
   AryTypePara[27].Other.S5Time := T#0MS;
   AryTypePara[27].Other."String" := '';
   AryTypePara[28].TypeName := '';
   AryTypePara[28].bit.Bit0 := FALSE;
   AryTypePara[28].bit.sp := 16#0000;
   AryTypePara[28].bit.Other.Bool_1 := FALSE;
   AryTypePara[28].bit.Other.Byte_2 := 16#00;
   AryTypePara[28].bit.Other.Int_1 := 0;
   AryTypePara[28].bit.Other."Char" := ' ';
   AryTypePara[28].Other.STxxxCCDProgNO := 0;
   AryTypePara[28].Other.FixtureEnable := FALSE;
   AryTypePara[28].Other.Byte_1 := 16#00;
   AryTypePara[28].Other.Int_1 := 0;
   AryTypePara[28].Other."Char" := ' ';
   AryTypePara[28].Other.Word_1 := 16#0000;
   AryTypePara[28].Other.DInt_1 := 0;
   AryTypePara[28].Other.DWord_1 := 16#0000_0000;
   AryTypePara[28].Other.Real_1 := 0.0;
   AryTypePara[28].Other.S5Time := T#0MS;
   AryTypePara[28].Other."String" := '';
   AryTypePara[29].TypeName := '';
   AryTypePara[29].bit.Bit0 := FALSE;
   AryTypePara[29].bit.sp := 16#0000;
   AryTypePara[29].bit.Other.Bool_1 := FALSE;
   AryTypePara[29].bit.Other.Byte_2 := 16#00;
   AryTypePara[29].bit.Other.Int_1 := 0;
   AryTypePara[29].bit.Other."Char" := ' ';
   AryTypePara[29].Other.STxxxCCDProgNO := 0;
   AryTypePara[29].Other.FixtureEnable := FALSE;
   AryTypePara[29].Other.Byte_1 := 16#00;
   AryTypePara[29].Other.Int_1 := 0;
   AryTypePara[29].Other."Char" := ' ';
   AryTypePara[29].Other.Word_1 := 16#0000;
   AryTypePara[29].Other.DInt_1 := 0;
   AryTypePara[29].Other.DWord_1 := 16#0000_0000;
   AryTypePara[29].Other.Real_1 := 0.0;
   AryTypePara[29].Other.S5Time := T#0MS;
   AryTypePara[29].Other."String" := '';
   AryTypePara[30].TypeName := '';
   AryTypePara[30].bit.Bit0 := FALSE;
   AryTypePara[30].bit.sp := 16#0000;
   AryTypePara[30].bit.Other.Bool_1 := FALSE;
   AryTypePara[30].bit.Other.Byte_2 := 16#00;
   AryTypePara[30].bit.Other.Int_1 := 0;
   AryTypePara[30].bit.Other."Char" := ' ';
   AryTypePara[30].Other.STxxxCCDProgNO := 0;
   AryTypePara[30].Other.FixtureEnable := FALSE;
   AryTypePara[30].Other.Byte_1 := 16#00;
   AryTypePara[30].Other.Int_1 := 0;
   AryTypePara[30].Other."Char" := ' ';
   AryTypePara[30].Other.Word_1 := 16#0000;
   AryTypePara[30].Other.DInt_1 := 0;
   AryTypePara[30].Other.DWord_1 := 16#0000_0000;
   AryTypePara[30].Other.Real_1 := 0.0;
   AryTypePara[30].Other.S5Time := T#0MS;
   AryTypePara[30].Other."String" := '';
   AryTypePara[31].TypeName := '';
   AryTypePara[31].bit.Bit0 := FALSE;
   AryTypePara[31].bit.sp := 16#0000;
   AryTypePara[31].bit.Other.Bool_1 := FALSE;
   AryTypePara[31].bit.Other.Byte_2 := 16#00;
   AryTypePara[31].bit.Other.Int_1 := 0;
   AryTypePara[31].bit.Other."Char" := ' ';
   AryTypePara[31].Other.STxxxCCDProgNO := 0;
   AryTypePara[31].Other.FixtureEnable := FALSE;
   AryTypePara[31].Other.Byte_1 := 16#00;
   AryTypePara[31].Other.Int_1 := 0;
   AryTypePara[31].Other."Char" := ' ';
   AryTypePara[31].Other.Word_1 := 16#0000;
   AryTypePara[31].Other.DInt_1 := 0;
   AryTypePara[31].Other.DWord_1 := 16#0000_0000;
   AryTypePara[31].Other.Real_1 := 0.0;
   AryTypePara[31].Other.S5Time := T#0MS;
   AryTypePara[31].Other."String" := '';
   AryTypePara[32].TypeName := '';
   AryTypePara[32].bit.Bit0 := FALSE;
   AryTypePara[32].bit.sp := 16#0000;
   AryTypePara[32].bit.Other.Bool_1 := FALSE;
   AryTypePara[32].bit.Other.Byte_2 := 16#00;
   AryTypePara[32].bit.Other.Int_1 := 0;
   AryTypePara[32].bit.Other."Char" := ' ';
   AryTypePara[32].Other.STxxxCCDProgNO := 0;
   AryTypePara[32].Other.FixtureEnable := FALSE;
   AryTypePara[32].Other.Byte_1 := 16#00;
   AryTypePara[32].Other.Int_1 := 0;
   AryTypePara[32].Other."Char" := ' ';
   AryTypePara[32].Other.Word_1 := 16#0000;
   AryTypePara[32].Other.DInt_1 := 0;
   AryTypePara[32].Other.DWord_1 := 16#0000_0000;
   AryTypePara[32].Other.Real_1 := 0.0;
   AryTypePara[32].Other.S5Time := T#0MS;
   AryTypePara[32].Other."String" := '';
   AryTypePara[33].TypeName := '';
   AryTypePara[33].bit.Bit0 := FALSE;
   AryTypePara[33].bit.sp := 16#0000;
   AryTypePara[33].bit.Other.Bool_1 := FALSE;
   AryTypePara[33].bit.Other.Byte_2 := 16#00;
   AryTypePara[33].bit.Other.Int_1 := 0;
   AryTypePara[33].bit.Other."Char" := ' ';
   AryTypePara[33].Other.STxxxCCDProgNO := 0;
   AryTypePara[33].Other.FixtureEnable := FALSE;
   AryTypePara[33].Other.Byte_1 := 16#00;
   AryTypePara[33].Other.Int_1 := 0;
   AryTypePara[33].Other."Char" := ' ';
   AryTypePara[33].Other.Word_1 := 16#0000;
   AryTypePara[33].Other.DInt_1 := 0;
   AryTypePara[33].Other.DWord_1 := 16#0000_0000;
   AryTypePara[33].Other.Real_1 := 0.0;
   AryTypePara[33].Other.S5Time := T#0MS;
   AryTypePara[33].Other."String" := '';
   AryTypePara[34].TypeName := '';
   AryTypePara[34].bit.Bit0 := FALSE;
   AryTypePara[34].bit.sp := 16#0000;
   AryTypePara[34].bit.Other.Bool_1 := FALSE;
   AryTypePara[34].bit.Other.Byte_2 := 16#00;
   AryTypePara[34].bit.Other.Int_1 := 0;
   AryTypePara[34].bit.Other."Char" := ' ';
   AryTypePara[34].Other.STxxxCCDProgNO := 0;
   AryTypePara[34].Other.FixtureEnable := FALSE;
   AryTypePara[34].Other.Byte_1 := 16#00;
   AryTypePara[34].Other.Int_1 := 0;
   AryTypePara[34].Other."Char" := ' ';
   AryTypePara[34].Other.Word_1 := 16#0000;
   AryTypePara[34].Other.DInt_1 := 0;
   AryTypePara[34].Other.DWord_1 := 16#0000_0000;
   AryTypePara[34].Other.Real_1 := 0.0;
   AryTypePara[34].Other.S5Time := T#0MS;
   AryTypePara[34].Other."String" := '';
   AryTypePara[35].TypeName := '';
   AryTypePara[35].bit.Bit0 := FALSE;
   AryTypePara[35].bit.sp := 16#0000;
   AryTypePara[35].bit.Other.Bool_1 := FALSE;
   AryTypePara[35].bit.Other.Byte_2 := 16#00;
   AryTypePara[35].bit.Other.Int_1 := 0;
   AryTypePara[35].bit.Other."Char" := ' ';
   AryTypePara[35].Other.STxxxCCDProgNO := 0;
   AryTypePara[35].Other.FixtureEnable := FALSE;
   AryTypePara[35].Other.Byte_1 := 16#00;
   AryTypePara[35].Other.Int_1 := 0;
   AryTypePara[35].Other."Char" := ' ';
   AryTypePara[35].Other.Word_1 := 16#0000;
   AryTypePara[35].Other.DInt_1 := 0;
   AryTypePara[35].Other.DWord_1 := 16#0000_0000;
   AryTypePara[35].Other.Real_1 := 0.0;
   AryTypePara[35].Other.S5Time := T#0MS;
   AryTypePara[35].Other."String" := '';
   AryTypePara[36].TypeName := '';
   AryTypePara[36].bit.Bit0 := FALSE;
   AryTypePara[36].bit.sp := 16#0000;
   AryTypePara[36].bit.Other.Bool_1 := FALSE;
   AryTypePara[36].bit.Other.Byte_2 := 16#00;
   AryTypePara[36].bit.Other.Int_1 := 0;
   AryTypePara[36].bit.Other."Char" := ' ';
   AryTypePara[36].Other.STxxxCCDProgNO := 0;
   AryTypePara[36].Other.FixtureEnable := FALSE;
   AryTypePara[36].Other.Byte_1 := 16#00;
   AryTypePara[36].Other.Int_1 := 0;
   AryTypePara[36].Other."Char" := ' ';
   AryTypePara[36].Other.Word_1 := 16#0000;
   AryTypePara[36].Other.DInt_1 := 0;
   AryTypePara[36].Other.DWord_1 := 16#0000_0000;
   AryTypePara[36].Other.Real_1 := 0.0;
   AryTypePara[36].Other.S5Time := T#0MS;
   AryTypePara[36].Other."String" := '';
   AryTypePara[37].TypeName := '';
   AryTypePara[37].bit.Bit0 := FALSE;
   AryTypePara[37].bit.sp := 16#0000;
   AryTypePara[37].bit.Other.Bool_1 := FALSE;
   AryTypePara[37].bit.Other.Byte_2 := 16#00;
   AryTypePara[37].bit.Other.Int_1 := 0;
   AryTypePara[37].bit.Other."Char" := ' ';
   AryTypePara[37].Other.STxxxCCDProgNO := 0;
   AryTypePara[37].Other.FixtureEnable := FALSE;
   AryTypePara[37].Other.Byte_1 := 16#00;
   AryTypePara[37].Other.Int_1 := 0;
   AryTypePara[37].Other."Char" := ' ';
   AryTypePara[37].Other.Word_1 := 16#0000;
   AryTypePara[37].Other.DInt_1 := 0;
   AryTypePara[37].Other.DWord_1 := 16#0000_0000;
   AryTypePara[37].Other.Real_1 := 0.0;
   AryTypePara[37].Other.S5Time := T#0MS;
   AryTypePara[37].Other."String" := '';
   AryTypePara[38].TypeName := '';
   AryTypePara[38].bit.Bit0 := FALSE;
   AryTypePara[38].bit.sp := 16#0000;
   AryTypePara[38].bit.Other.Bool_1 := FALSE;
   AryTypePara[38].bit.Other.Byte_2 := 16#00;
   AryTypePara[38].bit.Other.Int_1 := 0;
   AryTypePara[38].bit.Other."Char" := ' ';
   AryTypePara[38].Other.STxxxCCDProgNO := 0;
   AryTypePara[38].Other.FixtureEnable := FALSE;
   AryTypePara[38].Other.Byte_1 := 16#00;
   AryTypePara[38].Other.Int_1 := 0;
   AryTypePara[38].Other."Char" := ' ';
   AryTypePara[38].Other.Word_1 := 16#0000;
   AryTypePara[38].Other.DInt_1 := 0;
   AryTypePara[38].Other.DWord_1 := 16#0000_0000;
   AryTypePara[38].Other.Real_1 := 0.0;
   AryTypePara[38].Other.S5Time := T#0MS;
   AryTypePara[38].Other."String" := '';
   AryTypePara[39].TypeName := '';
   AryTypePara[39].bit.Bit0 := FALSE;
   AryTypePara[39].bit.sp := 16#0000;
   AryTypePara[39].bit.Other.Bool_1 := FALSE;
   AryTypePara[39].bit.Other.Byte_2 := 16#00;
   AryTypePara[39].bit.Other.Int_1 := 0;
   AryTypePara[39].bit.Other."Char" := ' ';
   AryTypePara[39].Other.STxxxCCDProgNO := 0;
   AryTypePara[39].Other.FixtureEnable := FALSE;
   AryTypePara[39].Other.Byte_1 := 16#00;
   AryTypePara[39].Other.Int_1 := 0;
   AryTypePara[39].Other."Char" := ' ';
   AryTypePara[39].Other.Word_1 := 16#0000;
   AryTypePara[39].Other.DInt_1 := 0;
   AryTypePara[39].Other.DWord_1 := 16#0000_0000;
   AryTypePara[39].Other.Real_1 := 0.0;
   AryTypePara[39].Other.S5Time := T#0MS;
   AryTypePara[39].Other."String" := '';
   AryTypePara[40].TypeName := '';
   AryTypePara[40].bit.Bit0 := FALSE;
   AryTypePara[40].bit.sp := 16#0000;
   AryTypePara[40].bit.Other.Bool_1 := FALSE;
   AryTypePara[40].bit.Other.Byte_2 := 16#00;
   AryTypePara[40].bit.Other.Int_1 := 0;
   AryTypePara[40].bit.Other."Char" := ' ';
   AryTypePara[40].Other.STxxxCCDProgNO := 0;
   AryTypePara[40].Other.FixtureEnable := FALSE;
   AryTypePara[40].Other.Byte_1 := 16#00;
   AryTypePara[40].Other.Int_1 := 0;
   AryTypePara[40].Other."Char" := ' ';
   AryTypePara[40].Other.Word_1 := 16#0000;
   AryTypePara[40].Other.DInt_1 := 0;
   AryTypePara[40].Other.DWord_1 := 16#0000_0000;
   AryTypePara[40].Other.Real_1 := 0.0;
   AryTypePara[40].Other.S5Time := T#0MS;
   AryTypePara[40].Other."String" := '';
   AryTypePara[41].TypeName := '';
   AryTypePara[41].bit.Bit0 := FALSE;
   AryTypePara[41].bit.sp := 16#0000;
   AryTypePara[41].bit.Other.Bool_1 := FALSE;
   AryTypePara[41].bit.Other.Byte_2 := 16#00;
   AryTypePara[41].bit.Other.Int_1 := 0;
   AryTypePara[41].bit.Other."Char" := ' ';
   AryTypePara[41].Other.STxxxCCDProgNO := 0;
   AryTypePara[41].Other.FixtureEnable := FALSE;
   AryTypePara[41].Other.Byte_1 := 16#00;
   AryTypePara[41].Other.Int_1 := 0;
   AryTypePara[41].Other."Char" := ' ';
   AryTypePara[41].Other.Word_1 := 16#0000;
   AryTypePara[41].Other.DInt_1 := 0;
   AryTypePara[41].Other.DWord_1 := 16#0000_0000;
   AryTypePara[41].Other.Real_1 := 0.0;
   AryTypePara[41].Other.S5Time := T#0MS;
   AryTypePara[41].Other."String" := '';
   AryTypePara[42].TypeName := '';
   AryTypePara[42].bit.Bit0 := FALSE;
   AryTypePara[42].bit.sp := 16#0000;
   AryTypePara[42].bit.Other.Bool_1 := FALSE;
   AryTypePara[42].bit.Other.Byte_2 := 16#00;
   AryTypePara[42].bit.Other.Int_1 := 0;
   AryTypePara[42].bit.Other."Char" := ' ';
   AryTypePara[42].Other.STxxxCCDProgNO := 0;
   AryTypePara[42].Other.FixtureEnable := FALSE;
   AryTypePara[42].Other.Byte_1 := 16#00;
   AryTypePara[42].Other.Int_1 := 0;
   AryTypePara[42].Other."Char" := ' ';
   AryTypePara[42].Other.Word_1 := 16#0000;
   AryTypePara[42].Other.DInt_1 := 0;
   AryTypePara[42].Other.DWord_1 := 16#0000_0000;
   AryTypePara[42].Other.Real_1 := 0.0;
   AryTypePara[42].Other.S5Time := T#0MS;
   AryTypePara[42].Other."String" := '';
   AryTypePara[43].TypeName := '';
   AryTypePara[43].bit.Bit0 := FALSE;
   AryTypePara[43].bit.sp := 16#0000;
   AryTypePara[43].bit.Other.Bool_1 := FALSE;
   AryTypePara[43].bit.Other.Byte_2 := 16#00;
   AryTypePara[43].bit.Other.Int_1 := 0;
   AryTypePara[43].bit.Other."Char" := ' ';
   AryTypePara[43].Other.STxxxCCDProgNO := 0;
   AryTypePara[43].Other.FixtureEnable := FALSE;
   AryTypePara[43].Other.Byte_1 := 16#00;
   AryTypePara[43].Other.Int_1 := 0;
   AryTypePara[43].Other."Char" := ' ';
   AryTypePara[43].Other.Word_1 := 16#0000;
   AryTypePara[43].Other.DInt_1 := 0;
   AryTypePara[43].Other.DWord_1 := 16#0000_0000;
   AryTypePara[43].Other.Real_1 := 0.0;
   AryTypePara[43].Other.S5Time := T#0MS;
   AryTypePara[43].Other."String" := '';
   AryTypePara[44].TypeName := '';
   AryTypePara[44].bit.Bit0 := FALSE;
   AryTypePara[44].bit.sp := 16#0000;
   AryTypePara[44].bit.Other.Bool_1 := FALSE;
   AryTypePara[44].bit.Other.Byte_2 := 16#00;
   AryTypePara[44].bit.Other.Int_1 := 0;
   AryTypePara[44].bit.Other."Char" := ' ';
   AryTypePara[44].Other.STxxxCCDProgNO := 0;
   AryTypePara[44].Other.FixtureEnable := FALSE;
   AryTypePara[44].Other.Byte_1 := 16#00;
   AryTypePara[44].Other.Int_1 := 0;
   AryTypePara[44].Other."Char" := ' ';
   AryTypePara[44].Other.Word_1 := 16#0000;
   AryTypePara[44].Other.DInt_1 := 0;
   AryTypePara[44].Other.DWord_1 := 16#0000_0000;
   AryTypePara[44].Other.Real_1 := 0.0;
   AryTypePara[44].Other.S5Time := T#0MS;
   AryTypePara[44].Other."String" := '';
   AryTypePara[45].TypeName := '';
   AryTypePara[45].bit.Bit0 := FALSE;
   AryTypePara[45].bit.sp := 16#0000;
   AryTypePara[45].bit.Other.Bool_1 := FALSE;
   AryTypePara[45].bit.Other.Byte_2 := 16#00;
   AryTypePara[45].bit.Other.Int_1 := 0;
   AryTypePara[45].bit.Other."Char" := ' ';
   AryTypePara[45].Other.STxxxCCDProgNO := 0;
   AryTypePara[45].Other.FixtureEnable := FALSE;
   AryTypePara[45].Other.Byte_1 := 16#00;
   AryTypePara[45].Other.Int_1 := 0;
   AryTypePara[45].Other."Char" := ' ';
   AryTypePara[45].Other.Word_1 := 16#0000;
   AryTypePara[45].Other.DInt_1 := 0;
   AryTypePara[45].Other.DWord_1 := 16#0000_0000;
   AryTypePara[45].Other.Real_1 := 0.0;
   AryTypePara[45].Other.S5Time := T#0MS;
   AryTypePara[45].Other."String" := '';
   AryTypePara[46].TypeName := '';
   AryTypePara[46].bit.Bit0 := FALSE;
   AryTypePara[46].bit.sp := 16#0000;
   AryTypePara[46].bit.Other.Bool_1 := FALSE;
   AryTypePara[46].bit.Other.Byte_2 := 16#00;
   AryTypePara[46].bit.Other.Int_1 := 0;
   AryTypePara[46].bit.Other."Char" := ' ';
   AryTypePara[46].Other.STxxxCCDProgNO := 0;
   AryTypePara[46].Other.FixtureEnable := FALSE;
   AryTypePara[46].Other.Byte_1 := 16#00;
   AryTypePara[46].Other.Int_1 := 0;
   AryTypePara[46].Other."Char" := ' ';
   AryTypePara[46].Other.Word_1 := 16#0000;
   AryTypePara[46].Other.DInt_1 := 0;
   AryTypePara[46].Other.DWord_1 := 16#0000_0000;
   AryTypePara[46].Other.Real_1 := 0.0;
   AryTypePara[46].Other.S5Time := T#0MS;
   AryTypePara[46].Other."String" := '';
   AryTypePara[47].TypeName := '';
   AryTypePara[47].bit.Bit0 := FALSE;
   AryTypePara[47].bit.sp := 16#0000;
   AryTypePara[47].bit.Other.Bool_1 := FALSE;
   AryTypePara[47].bit.Other.Byte_2 := 16#00;
   AryTypePara[47].bit.Other.Int_1 := 0;
   AryTypePara[47].bit.Other."Char" := ' ';
   AryTypePara[47].Other.STxxxCCDProgNO := 0;
   AryTypePara[47].Other.FixtureEnable := FALSE;
   AryTypePara[47].Other.Byte_1 := 16#00;
   AryTypePara[47].Other.Int_1 := 0;
   AryTypePara[47].Other."Char" := ' ';
   AryTypePara[47].Other.Word_1 := 16#0000;
   AryTypePara[47].Other.DInt_1 := 0;
   AryTypePara[47].Other.DWord_1 := 16#0000_0000;
   AryTypePara[47].Other.Real_1 := 0.0;
   AryTypePara[47].Other.S5Time := T#0MS;
   AryTypePara[47].Other."String" := '';
   AryTypePara[48].TypeName := '';
   AryTypePara[48].bit.Bit0 := FALSE;
   AryTypePara[48].bit.sp := 16#0000;
   AryTypePara[48].bit.Other.Bool_1 := FALSE;
   AryTypePara[48].bit.Other.Byte_2 := 16#00;
   AryTypePara[48].bit.Other.Int_1 := 0;
   AryTypePara[48].bit.Other."Char" := ' ';
   AryTypePara[48].Other.STxxxCCDProgNO := 0;
   AryTypePara[48].Other.FixtureEnable := FALSE;
   AryTypePara[48].Other.Byte_1 := 16#00;
   AryTypePara[48].Other.Int_1 := 0;
   AryTypePara[48].Other."Char" := ' ';
   AryTypePara[48].Other.Word_1 := 16#0000;
   AryTypePara[48].Other.DInt_1 := 0;
   AryTypePara[48].Other.DWord_1 := 16#0000_0000;
   AryTypePara[48].Other.Real_1 := 0.0;
   AryTypePara[48].Other.S5Time := T#0MS;
   AryTypePara[48].Other."String" := '';
   AryTypePara[49].TypeName := '';
   AryTypePara[49].bit.Bit0 := FALSE;
   AryTypePara[49].bit.sp := 16#0000;
   AryTypePara[49].bit.Other.Bool_1 := FALSE;
   AryTypePara[49].bit.Other.Byte_2 := 16#00;
   AryTypePara[49].bit.Other.Int_1 := 0;
   AryTypePara[49].bit.Other."Char" := ' ';
   AryTypePara[49].Other.STxxxCCDProgNO := 0;
   AryTypePara[49].Other.FixtureEnable := FALSE;
   AryTypePara[49].Other.Byte_1 := 16#00;
   AryTypePara[49].Other.Int_1 := 0;
   AryTypePara[49].Other."Char" := ' ';
   AryTypePara[49].Other.Word_1 := 16#0000;
   AryTypePara[49].Other.DInt_1 := 0;
   AryTypePara[49].Other.DWord_1 := 16#0000_0000;
   AryTypePara[49].Other.Real_1 := 0.0;
   AryTypePara[49].Other.S5Time := T#0MS;
   AryTypePara[49].Other."String" := '';
   AryTypePara[50].TypeName := '';
   AryTypePara[50].bit.Bit0 := FALSE;
   AryTypePara[50].bit.sp := 16#0000;
   AryTypePara[50].bit.Other.Bool_1 := FALSE;
   AryTypePara[50].bit.Other.Byte_2 := 16#00;
   AryTypePara[50].bit.Other.Int_1 := 0;
   AryTypePara[50].bit.Other."Char" := ' ';
   AryTypePara[50].Other.STxxxCCDProgNO := 0;
   AryTypePara[50].Other.FixtureEnable := FALSE;
   AryTypePara[50].Other.Byte_1 := 16#00;
   AryTypePara[50].Other.Int_1 := 0;
   AryTypePara[50].Other."Char" := ' ';
   AryTypePara[50].Other.Word_1 := 16#0000;
   AryTypePara[50].Other.DInt_1 := 0;
   AryTypePara[50].Other.DWord_1 := 16#0000_0000;
   AryTypePara[50].Other.Real_1 := 0.0;
   AryTypePara[50].Other.S5Time := T#0MS;
   AryTypePara[50].Other."String" := '';
   AryTypePara[51].TypeName := '';
   AryTypePara[51].bit.Bit0 := FALSE;
   AryTypePara[51].bit.sp := 16#0000;
   AryTypePara[51].bit.Other.Bool_1 := FALSE;
   AryTypePara[51].bit.Other.Byte_2 := 16#00;
   AryTypePara[51].bit.Other.Int_1 := 0;
   AryTypePara[51].bit.Other."Char" := ' ';
   AryTypePara[51].Other.STxxxCCDProgNO := 0;
   AryTypePara[51].Other.FixtureEnable := FALSE;
   AryTypePara[51].Other.Byte_1 := 16#00;
   AryTypePara[51].Other.Int_1 := 0;
   AryTypePara[51].Other."Char" := ' ';
   AryTypePara[51].Other.Word_1 := 16#0000;
   AryTypePara[51].Other.DInt_1 := 0;
   AryTypePara[51].Other.DWord_1 := 16#0000_0000;
   AryTypePara[51].Other.Real_1 := 0.0;
   AryTypePara[51].Other.S5Time := T#0MS;
   AryTypePara[51].Other."String" := '';
   AryTypePara[52].TypeName := '';
   AryTypePara[52].bit.Bit0 := FALSE;
   AryTypePara[52].bit.sp := 16#0000;
   AryTypePara[52].bit.Other.Bool_1 := FALSE;
   AryTypePara[52].bit.Other.Byte_2 := 16#00;
   AryTypePara[52].bit.Other.Int_1 := 0;
   AryTypePara[52].bit.Other."Char" := ' ';
   AryTypePara[52].Other.STxxxCCDProgNO := 0;
   AryTypePara[52].Other.FixtureEnable := FALSE;
   AryTypePara[52].Other.Byte_1 := 16#00;
   AryTypePara[52].Other.Int_1 := 0;
   AryTypePara[52].Other."Char" := ' ';
   AryTypePara[52].Other.Word_1 := 16#0000;
   AryTypePara[52].Other.DInt_1 := 0;
   AryTypePara[52].Other.DWord_1 := 16#0000_0000;
   AryTypePara[52].Other.Real_1 := 0.0;
   AryTypePara[52].Other.S5Time := T#0MS;
   AryTypePara[52].Other."String" := '';
   AryTypePara[53].TypeName := '';
   AryTypePara[53].bit.Bit0 := FALSE;
   AryTypePara[53].bit.sp := 16#0000;
   AryTypePara[53].bit.Other.Bool_1 := FALSE;
   AryTypePara[53].bit.Other.Byte_2 := 16#00;
   AryTypePara[53].bit.Other.Int_1 := 0;
   AryTypePara[53].bit.Other."Char" := ' ';
   AryTypePara[53].Other.STxxxCCDProgNO := 0;
   AryTypePara[53].Other.FixtureEnable := FALSE;
   AryTypePara[53].Other.Byte_1 := 16#00;
   AryTypePara[53].Other.Int_1 := 0;
   AryTypePara[53].Other."Char" := ' ';
   AryTypePara[53].Other.Word_1 := 16#0000;
   AryTypePara[53].Other.DInt_1 := 0;
   AryTypePara[53].Other.DWord_1 := 16#0000_0000;
   AryTypePara[53].Other.Real_1 := 0.0;
   AryTypePara[53].Other.S5Time := T#0MS;
   AryTypePara[53].Other."String" := '';
   AryTypePara[54].TypeName := '';
   AryTypePara[54].bit.Bit0 := FALSE;
   AryTypePara[54].bit.sp := 16#0000;
   AryTypePara[54].bit.Other.Bool_1 := FALSE;
   AryTypePara[54].bit.Other.Byte_2 := 16#00;
   AryTypePara[54].bit.Other.Int_1 := 0;
   AryTypePara[54].bit.Other."Char" := ' ';
   AryTypePara[54].Other.STxxxCCDProgNO := 0;
   AryTypePara[54].Other.FixtureEnable := FALSE;
   AryTypePara[54].Other.Byte_1 := 16#00;
   AryTypePara[54].Other.Int_1 := 0;
   AryTypePara[54].Other."Char" := ' ';
   AryTypePara[54].Other.Word_1 := 16#0000;
   AryTypePara[54].Other.DInt_1 := 0;
   AryTypePara[54].Other.DWord_1 := 16#0000_0000;
   AryTypePara[54].Other.Real_1 := 0.0;
   AryTypePara[54].Other.S5Time := T#0MS;
   AryTypePara[54].Other."String" := '';
   AryTypePara[55].TypeName := '';
   AryTypePara[55].bit.Bit0 := FALSE;
   AryTypePara[55].bit.sp := 16#0000;
   AryTypePara[55].bit.Other.Bool_1 := FALSE;
   AryTypePara[55].bit.Other.Byte_2 := 16#00;
   AryTypePara[55].bit.Other.Int_1 := 0;
   AryTypePara[55].bit.Other."Char" := ' ';
   AryTypePara[55].Other.STxxxCCDProgNO := 0;
   AryTypePara[55].Other.FixtureEnable := FALSE;
   AryTypePara[55].Other.Byte_1 := 16#00;
   AryTypePara[55].Other.Int_1 := 0;
   AryTypePara[55].Other."Char" := ' ';
   AryTypePara[55].Other.Word_1 := 16#0000;
   AryTypePara[55].Other.DInt_1 := 0;
   AryTypePara[55].Other.DWord_1 := 16#0000_0000;
   AryTypePara[55].Other.Real_1 := 0.0;
   AryTypePara[55].Other.S5Time := T#0MS;
   AryTypePara[55].Other."String" := '';
   AryTypePara[56].TypeName := '';
   AryTypePara[56].bit.Bit0 := FALSE;
   AryTypePara[56].bit.sp := 16#0000;
   AryTypePara[56].bit.Other.Bool_1 := FALSE;
   AryTypePara[56].bit.Other.Byte_2 := 16#00;
   AryTypePara[56].bit.Other.Int_1 := 0;
   AryTypePara[56].bit.Other."Char" := ' ';
   AryTypePara[56].Other.STxxxCCDProgNO := 0;
   AryTypePara[56].Other.FixtureEnable := FALSE;
   AryTypePara[56].Other.Byte_1 := 16#00;
   AryTypePara[56].Other.Int_1 := 0;
   AryTypePara[56].Other."Char" := ' ';
   AryTypePara[56].Other.Word_1 := 16#0000;
   AryTypePara[56].Other.DInt_1 := 0;
   AryTypePara[56].Other.DWord_1 := 16#0000_0000;
   AryTypePara[56].Other.Real_1 := 0.0;
   AryTypePara[56].Other.S5Time := T#0MS;
   AryTypePara[56].Other."String" := '';
   AryTypePara[57].TypeName := '';
   AryTypePara[57].bit.Bit0 := FALSE;
   AryTypePara[57].bit.sp := 16#0000;
   AryTypePara[57].bit.Other.Bool_1 := FALSE;
   AryTypePara[57].bit.Other.Byte_2 := 16#00;
   AryTypePara[57].bit.Other.Int_1 := 0;
   AryTypePara[57].bit.Other."Char" := ' ';
   AryTypePara[57].Other.STxxxCCDProgNO := 0;
   AryTypePara[57].Other.FixtureEnable := FALSE;
   AryTypePara[57].Other.Byte_1 := 16#00;
   AryTypePara[57].Other.Int_1 := 0;
   AryTypePara[57].Other."Char" := ' ';
   AryTypePara[57].Other.Word_1 := 16#0000;
   AryTypePara[57].Other.DInt_1 := 0;
   AryTypePara[57].Other.DWord_1 := 16#0000_0000;
   AryTypePara[57].Other.Real_1 := 0.0;
   AryTypePara[57].Other.S5Time := T#0MS;
   AryTypePara[57].Other."String" := '';
   AryTypePara[58].TypeName := '';
   AryTypePara[58].bit.Bit0 := FALSE;
   AryTypePara[58].bit.sp := 16#0000;
   AryTypePara[58].bit.Other.Bool_1 := FALSE;
   AryTypePara[58].bit.Other.Byte_2 := 16#00;
   AryTypePara[58].bit.Other.Int_1 := 0;
   AryTypePara[58].bit.Other."Char" := ' ';
   AryTypePara[58].Other.STxxxCCDProgNO := 0;
   AryTypePara[58].Other.FixtureEnable := FALSE;
   AryTypePara[58].Other.Byte_1 := 16#00;
   AryTypePara[58].Other.Int_1 := 0;
   AryTypePara[58].Other."Char" := ' ';
   AryTypePara[58].Other.Word_1 := 16#0000;
   AryTypePara[58].Other.DInt_1 := 0;
   AryTypePara[58].Other.DWord_1 := 16#0000_0000;
   AryTypePara[58].Other.Real_1 := 0.0;
   AryTypePara[58].Other.S5Time := T#0MS;
   AryTypePara[58].Other."String" := '';
   AryTypePara[59].TypeName := '';
   AryTypePara[59].bit.Bit0 := FALSE;
   AryTypePara[59].bit.sp := 16#0000;
   AryTypePara[59].bit.Other.Bool_1 := FALSE;
   AryTypePara[59].bit.Other.Byte_2 := 16#00;
   AryTypePara[59].bit.Other.Int_1 := 0;
   AryTypePara[59].bit.Other."Char" := ' ';
   AryTypePara[59].Other.STxxxCCDProgNO := 0;
   AryTypePara[59].Other.FixtureEnable := FALSE;
   AryTypePara[59].Other.Byte_1 := 16#00;
   AryTypePara[59].Other.Int_1 := 0;
   AryTypePara[59].Other."Char" := ' ';
   AryTypePara[59].Other.Word_1 := 16#0000;
   AryTypePara[59].Other.DInt_1 := 0;
   AryTypePara[59].Other.DWord_1 := 16#0000_0000;
   AryTypePara[59].Other.Real_1 := 0.0;
   AryTypePara[59].Other.S5Time := T#0MS;
   AryTypePara[59].Other."String" := '';
   AryTypePara[60].TypeName := '';
   AryTypePara[60].bit.Bit0 := FALSE;
   AryTypePara[60].bit.sp := 16#0000;
   AryTypePara[60].bit.Other.Bool_1 := FALSE;
   AryTypePara[60].bit.Other.Byte_2 := 16#00;
   AryTypePara[60].bit.Other.Int_1 := 0;
   AryTypePara[60].bit.Other."Char" := ' ';
   AryTypePara[60].Other.STxxxCCDProgNO := 0;
   AryTypePara[60].Other.FixtureEnable := FALSE;
   AryTypePara[60].Other.Byte_1 := 16#00;
   AryTypePara[60].Other.Int_1 := 0;
   AryTypePara[60].Other."Char" := ' ';
   AryTypePara[60].Other.Word_1 := 16#0000;
   AryTypePara[60].Other.DInt_1 := 0;
   AryTypePara[60].Other.DWord_1 := 16#0000_0000;
   AryTypePara[60].Other.Real_1 := 0.0;
   AryTypePara[60].Other.S5Time := T#0MS;
   AryTypePara[60].Other."String" := '';
   AryTypePara[61].TypeName := '';
   AryTypePara[61].bit.Bit0 := FALSE;
   AryTypePara[61].bit.sp := 16#0000;
   AryTypePara[61].bit.Other.Bool_1 := FALSE;
   AryTypePara[61].bit.Other.Byte_2 := 16#00;
   AryTypePara[61].bit.Other.Int_1 := 0;
   AryTypePara[61].bit.Other."Char" := ' ';
   AryTypePara[61].Other.STxxxCCDProgNO := 0;
   AryTypePara[61].Other.FixtureEnable := FALSE;
   AryTypePara[61].Other.Byte_1 := 16#00;
   AryTypePara[61].Other.Int_1 := 0;
   AryTypePara[61].Other."Char" := ' ';
   AryTypePara[61].Other.Word_1 := 16#0000;
   AryTypePara[61].Other.DInt_1 := 0;
   AryTypePara[61].Other.DWord_1 := 16#0000_0000;
   AryTypePara[61].Other.Real_1 := 0.0;
   AryTypePara[61].Other.S5Time := T#0MS;
   AryTypePara[61].Other."String" := '';
   AryTypePara[62].TypeName := '';
   AryTypePara[62].bit.Bit0 := FALSE;
   AryTypePara[62].bit.sp := 16#0000;
   AryTypePara[62].bit.Other.Bool_1 := FALSE;
   AryTypePara[62].bit.Other.Byte_2 := 16#00;
   AryTypePara[62].bit.Other.Int_1 := 0;
   AryTypePara[62].bit.Other."Char" := ' ';
   AryTypePara[62].Other.STxxxCCDProgNO := 0;
   AryTypePara[62].Other.FixtureEnable := FALSE;
   AryTypePara[62].Other.Byte_1 := 16#00;
   AryTypePara[62].Other.Int_1 := 0;
   AryTypePara[62].Other."Char" := ' ';
   AryTypePara[62].Other.Word_1 := 16#0000;
   AryTypePara[62].Other.DInt_1 := 0;
   AryTypePara[62].Other.DWord_1 := 16#0000_0000;
   AryTypePara[62].Other.Real_1 := 0.0;
   AryTypePara[62].Other.S5Time := T#0MS;
   AryTypePara[62].Other."String" := '';
   AryTypePara[63].TypeName := '';
   AryTypePara[63].bit.Bit0 := FALSE;
   AryTypePara[63].bit.sp := 16#0000;
   AryTypePara[63].bit.Other.Bool_1 := FALSE;
   AryTypePara[63].bit.Other.Byte_2 := 16#00;
   AryTypePara[63].bit.Other.Int_1 := 0;
   AryTypePara[63].bit.Other."Char" := ' ';
   AryTypePara[63].Other.STxxxCCDProgNO := 0;
   AryTypePara[63].Other.FixtureEnable := FALSE;
   AryTypePara[63].Other.Byte_1 := 16#00;
   AryTypePara[63].Other.Int_1 := 0;
   AryTypePara[63].Other."Char" := ' ';
   AryTypePara[63].Other.Word_1 := 16#0000;
   AryTypePara[63].Other.DInt_1 := 0;
   AryTypePara[63].Other.DWord_1 := 16#0000_0000;
   AryTypePara[63].Other.Real_1 := 0.0;
   AryTypePara[63].Other.S5Time := T#0MS;
   AryTypePara[63].Other."String" := '';
   AryTypePara[64].TypeName := '';
   AryTypePara[64].bit.Bit0 := FALSE;
   AryTypePara[64].bit.sp := 16#0000;
   AryTypePara[64].bit.Other.Bool_1 := FALSE;
   AryTypePara[64].bit.Other.Byte_2 := 16#00;
   AryTypePara[64].bit.Other.Int_1 := 0;
   AryTypePara[64].bit.Other."Char" := ' ';
   AryTypePara[64].Other.STxxxCCDProgNO := 0;
   AryTypePara[64].Other.FixtureEnable := FALSE;
   AryTypePara[64].Other.Byte_1 := 16#00;
   AryTypePara[64].Other.Int_1 := 0;
   AryTypePara[64].Other."Char" := ' ';
   AryTypePara[64].Other.Word_1 := 16#0000;
   AryTypePara[64].Other.DInt_1 := 0;
   AryTypePara[64].Other.DWord_1 := 16#0000_0000;
   AryTypePara[64].Other.Real_1 := 0.0;
   AryTypePara[64].Other.S5Time := T#0MS;
   AryTypePara[64].Other."String" := '';
   AryTypePara[65].TypeName := '';
   AryTypePara[65].bit.Bit0 := FALSE;
   AryTypePara[65].bit.sp := 16#0000;
   AryTypePara[65].bit.Other.Bool_1 := FALSE;
   AryTypePara[65].bit.Other.Byte_2 := 16#00;
   AryTypePara[65].bit.Other.Int_1 := 0;
   AryTypePara[65].bit.Other."Char" := ' ';
   AryTypePara[65].Other.STxxxCCDProgNO := 0;
   AryTypePara[65].Other.FixtureEnable := FALSE;
   AryTypePara[65].Other.Byte_1 := 16#00;
   AryTypePara[65].Other.Int_1 := 0;
   AryTypePara[65].Other."Char" := ' ';
   AryTypePara[65].Other.Word_1 := 16#0000;
   AryTypePara[65].Other.DInt_1 := 0;
   AryTypePara[65].Other.DWord_1 := 16#0000_0000;
   AryTypePara[65].Other.Real_1 := 0.0;
   AryTypePara[65].Other.S5Time := T#0MS;
   AryTypePara[65].Other."String" := '';
   AryTypePara[66].TypeName := '';
   AryTypePara[66].bit.Bit0 := FALSE;
   AryTypePara[66].bit.sp := 16#0000;
   AryTypePara[66].bit.Other.Bool_1 := FALSE;
   AryTypePara[66].bit.Other.Byte_2 := 16#00;
   AryTypePara[66].bit.Other.Int_1 := 0;
   AryTypePara[66].bit.Other."Char" := ' ';
   AryTypePara[66].Other.STxxxCCDProgNO := 0;
   AryTypePara[66].Other.FixtureEnable := FALSE;
   AryTypePara[66].Other.Byte_1 := 16#00;
   AryTypePara[66].Other.Int_1 := 0;
   AryTypePara[66].Other."Char" := ' ';
   AryTypePara[66].Other.Word_1 := 16#0000;
   AryTypePara[66].Other.DInt_1 := 0;
   AryTypePara[66].Other.DWord_1 := 16#0000_0000;
   AryTypePara[66].Other.Real_1 := 0.0;
   AryTypePara[66].Other.S5Time := T#0MS;
   AryTypePara[66].Other."String" := '';
   AryTypePara[67].TypeName := '';
   AryTypePara[67].bit.Bit0 := FALSE;
   AryTypePara[67].bit.sp := 16#0000;
   AryTypePara[67].bit.Other.Bool_1 := FALSE;
   AryTypePara[67].bit.Other.Byte_2 := 16#00;
   AryTypePara[67].bit.Other.Int_1 := 0;
   AryTypePara[67].bit.Other."Char" := ' ';
   AryTypePara[67].Other.STxxxCCDProgNO := 0;
   AryTypePara[67].Other.FixtureEnable := FALSE;
   AryTypePara[67].Other.Byte_1 := 16#00;
   AryTypePara[67].Other.Int_1 := 0;
   AryTypePara[67].Other."Char" := ' ';
   AryTypePara[67].Other.Word_1 := 16#0000;
   AryTypePara[67].Other.DInt_1 := 0;
   AryTypePara[67].Other.DWord_1 := 16#0000_0000;
   AryTypePara[67].Other.Real_1 := 0.0;
   AryTypePara[67].Other.S5Time := T#0MS;
   AryTypePara[67].Other."String" := '';
   AryTypePara[68].TypeName := '';
   AryTypePara[68].bit.Bit0 := FALSE;
   AryTypePara[68].bit.sp := 16#0000;
   AryTypePara[68].bit.Other.Bool_1 := FALSE;
   AryTypePara[68].bit.Other.Byte_2 := 16#00;
   AryTypePara[68].bit.Other.Int_1 := 0;
   AryTypePara[68].bit.Other."Char" := ' ';
   AryTypePara[68].Other.STxxxCCDProgNO := 0;
   AryTypePara[68].Other.FixtureEnable := FALSE;
   AryTypePara[68].Other.Byte_1 := 16#00;
   AryTypePara[68].Other.Int_1 := 0;
   AryTypePara[68].Other."Char" := ' ';
   AryTypePara[68].Other.Word_1 := 16#0000;
   AryTypePara[68].Other.DInt_1 := 0;
   AryTypePara[68].Other.DWord_1 := 16#0000_0000;
   AryTypePara[68].Other.Real_1 := 0.0;
   AryTypePara[68].Other.S5Time := T#0MS;
   AryTypePara[68].Other."String" := '';
   AryTypePara[69].TypeName := '';
   AryTypePara[69].bit.Bit0 := FALSE;
   AryTypePara[69].bit.sp := 16#0000;
   AryTypePara[69].bit.Other.Bool_1 := FALSE;
   AryTypePara[69].bit.Other.Byte_2 := 16#00;
   AryTypePara[69].bit.Other.Int_1 := 0;
   AryTypePara[69].bit.Other."Char" := ' ';
   AryTypePara[69].Other.STxxxCCDProgNO := 0;
   AryTypePara[69].Other.FixtureEnable := FALSE;
   AryTypePara[69].Other.Byte_1 := 16#00;
   AryTypePara[69].Other.Int_1 := 0;
   AryTypePara[69].Other."Char" := ' ';
   AryTypePara[69].Other.Word_1 := 16#0000;
   AryTypePara[69].Other.DInt_1 := 0;
   AryTypePara[69].Other.DWord_1 := 16#0000_0000;
   AryTypePara[69].Other.Real_1 := 0.0;
   AryTypePara[69].Other.S5Time := T#0MS;
   AryTypePara[69].Other."String" := '';
   AryTypePara[70].TypeName := '';
   AryTypePara[70].bit.Bit0 := FALSE;
   AryTypePara[70].bit.sp := 16#0000;
   AryTypePara[70].bit.Other.Bool_1 := FALSE;
   AryTypePara[70].bit.Other.Byte_2 := 16#00;
   AryTypePara[70].bit.Other.Int_1 := 0;
   AryTypePara[70].bit.Other."Char" := ' ';
   AryTypePara[70].Other.STxxxCCDProgNO := 0;
   AryTypePara[70].Other.FixtureEnable := FALSE;
   AryTypePara[70].Other.Byte_1 := 16#00;
   AryTypePara[70].Other.Int_1 := 0;
   AryTypePara[70].Other."Char" := ' ';
   AryTypePara[70].Other.Word_1 := 16#0000;
   AryTypePara[70].Other.DInt_1 := 0;
   AryTypePara[70].Other.DWord_1 := 16#0000_0000;
   AryTypePara[70].Other.Real_1 := 0.0;
   AryTypePara[70].Other.S5Time := T#0MS;
   AryTypePara[70].Other."String" := '';
   AryTypePara[71].TypeName := '';
   AryTypePara[71].bit.Bit0 := FALSE;
   AryTypePara[71].bit.sp := 16#0000;
   AryTypePara[71].bit.Other.Bool_1 := FALSE;
   AryTypePara[71].bit.Other.Byte_2 := 16#00;
   AryTypePara[71].bit.Other.Int_1 := 0;
   AryTypePara[71].bit.Other."Char" := ' ';
   AryTypePara[71].Other.STxxxCCDProgNO := 0;
   AryTypePara[71].Other.FixtureEnable := FALSE;
   AryTypePara[71].Other.Byte_1 := 16#00;
   AryTypePara[71].Other.Int_1 := 0;
   AryTypePara[71].Other."Char" := ' ';
   AryTypePara[71].Other.Word_1 := 16#0000;
   AryTypePara[71].Other.DInt_1 := 0;
   AryTypePara[71].Other.DWord_1 := 16#0000_0000;
   AryTypePara[71].Other.Real_1 := 0.0;
   AryTypePara[71].Other.S5Time := T#0MS;
   AryTypePara[71].Other."String" := '';
   AryTypePara[72].TypeName := '';
   AryTypePara[72].bit.Bit0 := FALSE;
   AryTypePara[72].bit.sp := 16#0000;
   AryTypePara[72].bit.Other.Bool_1 := FALSE;
   AryTypePara[72].bit.Other.Byte_2 := 16#00;
   AryTypePara[72].bit.Other.Int_1 := 0;
   AryTypePara[72].bit.Other."Char" := ' ';
   AryTypePara[72].Other.STxxxCCDProgNO := 0;
   AryTypePara[72].Other.FixtureEnable := FALSE;
   AryTypePara[72].Other.Byte_1 := 16#00;
   AryTypePara[72].Other.Int_1 := 0;
   AryTypePara[72].Other."Char" := ' ';
   AryTypePara[72].Other.Word_1 := 16#0000;
   AryTypePara[72].Other.DInt_1 := 0;
   AryTypePara[72].Other.DWord_1 := 16#0000_0000;
   AryTypePara[72].Other.Real_1 := 0.0;
   AryTypePara[72].Other.S5Time := T#0MS;
   AryTypePara[72].Other."String" := '';
   AryTypePara[73].TypeName := '';
   AryTypePara[73].bit.Bit0 := FALSE;
   AryTypePara[73].bit.sp := 16#0000;
   AryTypePara[73].bit.Other.Bool_1 := FALSE;
   AryTypePara[73].bit.Other.Byte_2 := 16#00;
   AryTypePara[73].bit.Other.Int_1 := 0;
   AryTypePara[73].bit.Other."Char" := ' ';
   AryTypePara[73].Other.STxxxCCDProgNO := 0;
   AryTypePara[73].Other.FixtureEnable := FALSE;
   AryTypePara[73].Other.Byte_1 := 16#00;
   AryTypePara[73].Other.Int_1 := 0;
   AryTypePara[73].Other."Char" := ' ';
   AryTypePara[73].Other.Word_1 := 16#0000;
   AryTypePara[73].Other.DInt_1 := 0;
   AryTypePara[73].Other.DWord_1 := 16#0000_0000;
   AryTypePara[73].Other.Real_1 := 0.0;
   AryTypePara[73].Other.S5Time := T#0MS;
   AryTypePara[73].Other."String" := '';
   AryTypePara[74].TypeName := '';
   AryTypePara[74].bit.Bit0 := FALSE;
   AryTypePara[74].bit.sp := 16#0000;
   AryTypePara[74].bit.Other.Bool_1 := FALSE;
   AryTypePara[74].bit.Other.Byte_2 := 16#00;
   AryTypePara[74].bit.Other.Int_1 := 0;
   AryTypePara[74].bit.Other."Char" := ' ';
   AryTypePara[74].Other.STxxxCCDProgNO := 0;
   AryTypePara[74].Other.FixtureEnable := FALSE;
   AryTypePara[74].Other.Byte_1 := 16#00;
   AryTypePara[74].Other.Int_1 := 0;
   AryTypePara[74].Other."Char" := ' ';
   AryTypePara[74].Other.Word_1 := 16#0000;
   AryTypePara[74].Other.DInt_1 := 0;
   AryTypePara[74].Other.DWord_1 := 16#0000_0000;
   AryTypePara[74].Other.Real_1 := 0.0;
   AryTypePara[74].Other.S5Time := T#0MS;
   AryTypePara[74].Other."String" := '';
   AryTypePara[75].TypeName := '';
   AryTypePara[75].bit.Bit0 := FALSE;
   AryTypePara[75].bit.sp := 16#0000;
   AryTypePara[75].bit.Other.Bool_1 := FALSE;
   AryTypePara[75].bit.Other.Byte_2 := 16#00;
   AryTypePara[75].bit.Other.Int_1 := 0;
   AryTypePara[75].bit.Other."Char" := ' ';
   AryTypePara[75].Other.STxxxCCDProgNO := 0;
   AryTypePara[75].Other.FixtureEnable := FALSE;
   AryTypePara[75].Other.Byte_1 := 16#00;
   AryTypePara[75].Other.Int_1 := 0;
   AryTypePara[75].Other."Char" := ' ';
   AryTypePara[75].Other.Word_1 := 16#0000;
   AryTypePara[75].Other.DInt_1 := 0;
   AryTypePara[75].Other.DWord_1 := 16#0000_0000;
   AryTypePara[75].Other.Real_1 := 0.0;
   AryTypePara[75].Other.S5Time := T#0MS;
   AryTypePara[75].Other."String" := '';
   AryTypePara[76].TypeName := '';
   AryTypePara[76].bit.Bit0 := FALSE;
   AryTypePara[76].bit.sp := 16#0000;
   AryTypePara[76].bit.Other.Bool_1 := FALSE;
   AryTypePara[76].bit.Other.Byte_2 := 16#00;
   AryTypePara[76].bit.Other.Int_1 := 0;
   AryTypePara[76].bit.Other."Char" := ' ';
   AryTypePara[76].Other.STxxxCCDProgNO := 0;
   AryTypePara[76].Other.FixtureEnable := FALSE;
   AryTypePara[76].Other.Byte_1 := 16#00;
   AryTypePara[76].Other.Int_1 := 0;
   AryTypePara[76].Other."Char" := ' ';
   AryTypePara[76].Other.Word_1 := 16#0000;
   AryTypePara[76].Other.DInt_1 := 0;
   AryTypePara[76].Other.DWord_1 := 16#0000_0000;
   AryTypePara[76].Other.Real_1 := 0.0;
   AryTypePara[76].Other.S5Time := T#0MS;
   AryTypePara[76].Other."String" := '';
   AryTypePara[77].TypeName := '';
   AryTypePara[77].bit.Bit0 := FALSE;
   AryTypePara[77].bit.sp := 16#0000;
   AryTypePara[77].bit.Other.Bool_1 := FALSE;
   AryTypePara[77].bit.Other.Byte_2 := 16#00;
   AryTypePara[77].bit.Other.Int_1 := 0;
   AryTypePara[77].bit.Other."Char" := ' ';
   AryTypePara[77].Other.STxxxCCDProgNO := 0;
   AryTypePara[77].Other.FixtureEnable := FALSE;
   AryTypePara[77].Other.Byte_1 := 16#00;
   AryTypePara[77].Other.Int_1 := 0;
   AryTypePara[77].Other."Char" := ' ';
   AryTypePara[77].Other.Word_1 := 16#0000;
   AryTypePara[77].Other.DInt_1 := 0;
   AryTypePara[77].Other.DWord_1 := 16#0000_0000;
   AryTypePara[77].Other.Real_1 := 0.0;
   AryTypePara[77].Other.S5Time := T#0MS;
   AryTypePara[77].Other."String" := '';
   AryTypePara[78].TypeName := '';
   AryTypePara[78].bit.Bit0 := FALSE;
   AryTypePara[78].bit.sp := 16#0000;
   AryTypePara[78].bit.Other.Bool_1 := FALSE;
   AryTypePara[78].bit.Other.Byte_2 := 16#00;
   AryTypePara[78].bit.Other.Int_1 := 0;
   AryTypePara[78].bit.Other."Char" := ' ';
   AryTypePara[78].Other.STxxxCCDProgNO := 0;
   AryTypePara[78].Other.FixtureEnable := FALSE;
   AryTypePara[78].Other.Byte_1 := 16#00;
   AryTypePara[78].Other.Int_1 := 0;
   AryTypePara[78].Other."Char" := ' ';
   AryTypePara[78].Other.Word_1 := 16#0000;
   AryTypePara[78].Other.DInt_1 := 0;
   AryTypePara[78].Other.DWord_1 := 16#0000_0000;
   AryTypePara[78].Other.Real_1 := 0.0;
   AryTypePara[78].Other.S5Time := T#0MS;
   AryTypePara[78].Other."String" := '';
   AryTypePara[79].TypeName := '';
   AryTypePara[79].bit.Bit0 := FALSE;
   AryTypePara[79].bit.sp := 16#0000;
   AryTypePara[79].bit.Other.Bool_1 := FALSE;
   AryTypePara[79].bit.Other.Byte_2 := 16#00;
   AryTypePara[79].bit.Other.Int_1 := 0;
   AryTypePara[79].bit.Other."Char" := ' ';
   AryTypePara[79].Other.STxxxCCDProgNO := 0;
   AryTypePara[79].Other.FixtureEnable := FALSE;
   AryTypePara[79].Other.Byte_1 := 16#00;
   AryTypePara[79].Other.Int_1 := 0;
   AryTypePara[79].Other."Char" := ' ';
   AryTypePara[79].Other.Word_1 := 16#0000;
   AryTypePara[79].Other.DInt_1 := 0;
   AryTypePara[79].Other.DWord_1 := 16#0000_0000;
   AryTypePara[79].Other.Real_1 := 0.0;
   AryTypePara[79].Other.S5Time := T#0MS;
   AryTypePara[79].Other."String" := '';
   AryTypePara[80].TypeName := '';
   AryTypePara[80].bit.Bit0 := FALSE;
   AryTypePara[80].bit.sp := 16#0000;
   AryTypePara[80].bit.Other.Bool_1 := FALSE;
   AryTypePara[80].bit.Other.Byte_2 := 16#00;
   AryTypePara[80].bit.Other.Int_1 := 0;
   AryTypePara[80].bit.Other."Char" := ' ';
   AryTypePara[80].Other.STxxxCCDProgNO := 0;
   AryTypePara[80].Other.FixtureEnable := FALSE;
   AryTypePara[80].Other.Byte_1 := 16#00;
   AryTypePara[80].Other.Int_1 := 0;
   AryTypePara[80].Other."Char" := ' ';
   AryTypePara[80].Other.Word_1 := 16#0000;
   AryTypePara[80].Other.DInt_1 := 0;
   AryTypePara[80].Other.DWord_1 := 16#0000_0000;
   AryTypePara[80].Other.Real_1 := 0.0;
   AryTypePara[80].Other.S5Time := T#0MS;
   AryTypePara[80].Other."String" := '';
   AryTypePara[81].TypeName := '';
   AryTypePara[81].bit.Bit0 := FALSE;
   AryTypePara[81].bit.sp := 16#0000;
   AryTypePara[81].bit.Other.Bool_1 := FALSE;
   AryTypePara[81].bit.Other.Byte_2 := 16#00;
   AryTypePara[81].bit.Other.Int_1 := 0;
   AryTypePara[81].bit.Other."Char" := ' ';
   AryTypePara[81].Other.STxxxCCDProgNO := 0;
   AryTypePara[81].Other.FixtureEnable := FALSE;
   AryTypePara[81].Other.Byte_1 := 16#00;
   AryTypePara[81].Other.Int_1 := 0;
   AryTypePara[81].Other."Char" := ' ';
   AryTypePara[81].Other.Word_1 := 16#0000;
   AryTypePara[81].Other.DInt_1 := 0;
   AryTypePara[81].Other.DWord_1 := 16#0000_0000;
   AryTypePara[81].Other.Real_1 := 0.0;
   AryTypePara[81].Other.S5Time := T#0MS;
   AryTypePara[81].Other."String" := '';
   AryTypePara[82].TypeName := '';
   AryTypePara[82].bit.Bit0 := FALSE;
   AryTypePara[82].bit.sp := 16#0000;
   AryTypePara[82].bit.Other.Bool_1 := FALSE;
   AryTypePara[82].bit.Other.Byte_2 := 16#00;
   AryTypePara[82].bit.Other.Int_1 := 0;
   AryTypePara[82].bit.Other."Char" := ' ';
   AryTypePara[82].Other.STxxxCCDProgNO := 0;
   AryTypePara[82].Other.FixtureEnable := FALSE;
   AryTypePara[82].Other.Byte_1 := 16#00;
   AryTypePara[82].Other.Int_1 := 0;
   AryTypePara[82].Other."Char" := ' ';
   AryTypePara[82].Other.Word_1 := 16#0000;
   AryTypePara[82].Other.DInt_1 := 0;
   AryTypePara[82].Other.DWord_1 := 16#0000_0000;
   AryTypePara[82].Other.Real_1 := 0.0;
   AryTypePara[82].Other.S5Time := T#0MS;
   AryTypePara[82].Other."String" := '';
   AryTypePara[83].TypeName := '';
   AryTypePara[83].bit.Bit0 := FALSE;
   AryTypePara[83].bit.sp := 16#0000;
   AryTypePara[83].bit.Other.Bool_1 := FALSE;
   AryTypePara[83].bit.Other.Byte_2 := 16#00;
   AryTypePara[83].bit.Other.Int_1 := 0;
   AryTypePara[83].bit.Other."Char" := ' ';
   AryTypePara[83].Other.STxxxCCDProgNO := 0;
   AryTypePara[83].Other.FixtureEnable := FALSE;
   AryTypePara[83].Other.Byte_1 := 16#00;
   AryTypePara[83].Other.Int_1 := 0;
   AryTypePara[83].Other."Char" := ' ';
   AryTypePara[83].Other.Word_1 := 16#0000;
   AryTypePara[83].Other.DInt_1 := 0;
   AryTypePara[83].Other.DWord_1 := 16#0000_0000;
   AryTypePara[83].Other.Real_1 := 0.0;
   AryTypePara[83].Other.S5Time := T#0MS;
   AryTypePara[83].Other."String" := '';
   AryTypePara[84].TypeName := '';
   AryTypePara[84].bit.Bit0 := FALSE;
   AryTypePara[84].bit.sp := 16#0000;
   AryTypePara[84].bit.Other.Bool_1 := FALSE;
   AryTypePara[84].bit.Other.Byte_2 := 16#00;
   AryTypePara[84].bit.Other.Int_1 := 0;
   AryTypePara[84].bit.Other."Char" := ' ';
   AryTypePara[84].Other.STxxxCCDProgNO := 0;
   AryTypePara[84].Other.FixtureEnable := FALSE;
   AryTypePara[84].Other.Byte_1 := 16#00;
   AryTypePara[84].Other.Int_1 := 0;
   AryTypePara[84].Other."Char" := ' ';
   AryTypePara[84].Other.Word_1 := 16#0000;
   AryTypePara[84].Other.DInt_1 := 0;
   AryTypePara[84].Other.DWord_1 := 16#0000_0000;
   AryTypePara[84].Other.Real_1 := 0.0;
   AryTypePara[84].Other.S5Time := T#0MS;
   AryTypePara[84].Other."String" := '';
   AryTypePara[85].TypeName := '';
   AryTypePara[85].bit.Bit0 := FALSE;
   AryTypePara[85].bit.sp := 16#0000;
   AryTypePara[85].bit.Other.Bool_1 := FALSE;
   AryTypePara[85].bit.Other.Byte_2 := 16#00;
   AryTypePara[85].bit.Other.Int_1 := 0;
   AryTypePara[85].bit.Other."Char" := ' ';
   AryTypePara[85].Other.STxxxCCDProgNO := 0;
   AryTypePara[85].Other.FixtureEnable := FALSE;
   AryTypePara[85].Other.Byte_1 := 16#00;
   AryTypePara[85].Other.Int_1 := 0;
   AryTypePara[85].Other."Char" := ' ';
   AryTypePara[85].Other.Word_1 := 16#0000;
   AryTypePara[85].Other.DInt_1 := 0;
   AryTypePara[85].Other.DWord_1 := 16#0000_0000;
   AryTypePara[85].Other.Real_1 := 0.0;
   AryTypePara[85].Other.S5Time := T#0MS;
   AryTypePara[85].Other."String" := '';
   AryTypePara[86].TypeName := '';
   AryTypePara[86].bit.Bit0 := FALSE;
   AryTypePara[86].bit.sp := 16#0000;
   AryTypePara[86].bit.Other.Bool_1 := FALSE;
   AryTypePara[86].bit.Other.Byte_2 := 16#00;
   AryTypePara[86].bit.Other.Int_1 := 0;
   AryTypePara[86].bit.Other."Char" := ' ';
   AryTypePara[86].Other.STxxxCCDProgNO := 0;
   AryTypePara[86].Other.FixtureEnable := FALSE;
   AryTypePara[86].Other.Byte_1 := 16#00;
   AryTypePara[86].Other.Int_1 := 0;
   AryTypePara[86].Other."Char" := ' ';
   AryTypePara[86].Other.Word_1 := 16#0000;
   AryTypePara[86].Other.DInt_1 := 0;
   AryTypePara[86].Other.DWord_1 := 16#0000_0000;
   AryTypePara[86].Other.Real_1 := 0.0;
   AryTypePara[86].Other.S5Time := T#0MS;
   AryTypePara[86].Other."String" := '';
   AryTypePara[87].TypeName := '';
   AryTypePara[87].bit.Bit0 := FALSE;
   AryTypePara[87].bit.sp := 16#0000;
   AryTypePara[87].bit.Other.Bool_1 := FALSE;
   AryTypePara[87].bit.Other.Byte_2 := 16#00;
   AryTypePara[87].bit.Other.Int_1 := 0;
   AryTypePara[87].bit.Other."Char" := ' ';
   AryTypePara[87].Other.STxxxCCDProgNO := 0;
   AryTypePara[87].Other.FixtureEnable := FALSE;
   AryTypePara[87].Other.Byte_1 := 16#00;
   AryTypePara[87].Other.Int_1 := 0;
   AryTypePara[87].Other."Char" := ' ';
   AryTypePara[87].Other.Word_1 := 16#0000;
   AryTypePara[87].Other.DInt_1 := 0;
   AryTypePara[87].Other.DWord_1 := 16#0000_0000;
   AryTypePara[87].Other.Real_1 := 0.0;
   AryTypePara[87].Other.S5Time := T#0MS;
   AryTypePara[87].Other."String" := '';
   AryTypePara[88].TypeName := '';
   AryTypePara[88].bit.Bit0 := FALSE;
   AryTypePara[88].bit.sp := 16#0000;
   AryTypePara[88].bit.Other.Bool_1 := FALSE;
   AryTypePara[88].bit.Other.Byte_2 := 16#00;
   AryTypePara[88].bit.Other.Int_1 := 0;
   AryTypePara[88].bit.Other."Char" := ' ';
   AryTypePara[88].Other.STxxxCCDProgNO := 0;
   AryTypePara[88].Other.FixtureEnable := FALSE;
   AryTypePara[88].Other.Byte_1 := 16#00;
   AryTypePara[88].Other.Int_1 := 0;
   AryTypePara[88].Other."Char" := ' ';
   AryTypePara[88].Other.Word_1 := 16#0000;
   AryTypePara[88].Other.DInt_1 := 0;
   AryTypePara[88].Other.DWord_1 := 16#0000_0000;
   AryTypePara[88].Other.Real_1 := 0.0;
   AryTypePara[88].Other.S5Time := T#0MS;
   AryTypePara[88].Other."String" := '';
   AryTypePara[89].TypeName := '';
   AryTypePara[89].bit.Bit0 := FALSE;
   AryTypePara[89].bit.sp := 16#0000;
   AryTypePara[89].bit.Other.Bool_1 := FALSE;
   AryTypePara[89].bit.Other.Byte_2 := 16#00;
   AryTypePara[89].bit.Other.Int_1 := 0;
   AryTypePara[89].bit.Other."Char" := ' ';
   AryTypePara[89].Other.STxxxCCDProgNO := 0;
   AryTypePara[89].Other.FixtureEnable := FALSE;
   AryTypePara[89].Other.Byte_1 := 16#00;
   AryTypePara[89].Other.Int_1 := 0;
   AryTypePara[89].Other."Char" := ' ';
   AryTypePara[89].Other.Word_1 := 16#0000;
   AryTypePara[89].Other.DInt_1 := 0;
   AryTypePara[89].Other.DWord_1 := 16#0000_0000;
   AryTypePara[89].Other.Real_1 := 0.0;
   AryTypePara[89].Other.S5Time := T#0MS;
   AryTypePara[89].Other."String" := '';
   AryTypePara[90].TypeName := '';
   AryTypePara[90].bit.Bit0 := FALSE;
   AryTypePara[90].bit.sp := 16#0000;
   AryTypePara[90].bit.Other.Bool_1 := FALSE;
   AryTypePara[90].bit.Other.Byte_2 := 16#00;
   AryTypePara[90].bit.Other.Int_1 := 0;
   AryTypePara[90].bit.Other."Char" := ' ';
   AryTypePara[90].Other.STxxxCCDProgNO := 0;
   AryTypePara[90].Other.FixtureEnable := FALSE;
   AryTypePara[90].Other.Byte_1 := 16#00;
   AryTypePara[90].Other.Int_1 := 0;
   AryTypePara[90].Other."Char" := ' ';
   AryTypePara[90].Other.Word_1 := 16#0000;
   AryTypePara[90].Other.DInt_1 := 0;
   AryTypePara[90].Other.DWord_1 := 16#0000_0000;
   AryTypePara[90].Other.Real_1 := 0.0;
   AryTypePara[90].Other.S5Time := T#0MS;
   AryTypePara[90].Other."String" := '';
   AryTypePara[91].TypeName := '';
   AryTypePara[91].bit.Bit0 := FALSE;
   AryTypePara[91].bit.sp := 16#0000;
   AryTypePara[91].bit.Other.Bool_1 := FALSE;
   AryTypePara[91].bit.Other.Byte_2 := 16#00;
   AryTypePara[91].bit.Other.Int_1 := 0;
   AryTypePara[91].bit.Other."Char" := ' ';
   AryTypePara[91].Other.STxxxCCDProgNO := 0;
   AryTypePara[91].Other.FixtureEnable := FALSE;
   AryTypePara[91].Other.Byte_1 := 16#00;
   AryTypePara[91].Other.Int_1 := 0;
   AryTypePara[91].Other."Char" := ' ';
   AryTypePara[91].Other.Word_1 := 16#0000;
   AryTypePara[91].Other.DInt_1 := 0;
   AryTypePara[91].Other.DWord_1 := 16#0000_0000;
   AryTypePara[91].Other.Real_1 := 0.0;
   AryTypePara[91].Other.S5Time := T#0MS;
   AryTypePara[91].Other."String" := '';
   AryTypePara[92].TypeName := '';
   AryTypePara[92].bit.Bit0 := FALSE;
   AryTypePara[92].bit.sp := 16#0000;
   AryTypePara[92].bit.Other.Bool_1 := FALSE;
   AryTypePara[92].bit.Other.Byte_2 := 16#00;
   AryTypePara[92].bit.Other.Int_1 := 0;
   AryTypePara[92].bit.Other."Char" := ' ';
   AryTypePara[92].Other.STxxxCCDProgNO := 0;
   AryTypePara[92].Other.FixtureEnable := FALSE;
   AryTypePara[92].Other.Byte_1 := 16#00;
   AryTypePara[92].Other.Int_1 := 0;
   AryTypePara[92].Other."Char" := ' ';
   AryTypePara[92].Other.Word_1 := 16#0000;
   AryTypePara[92].Other.DInt_1 := 0;
   AryTypePara[92].Other.DWord_1 := 16#0000_0000;
   AryTypePara[92].Other.Real_1 := 0.0;
   AryTypePara[92].Other.S5Time := T#0MS;
   AryTypePara[92].Other."String" := '';
   AryTypePara[93].TypeName := '';
   AryTypePara[93].bit.Bit0 := FALSE;
   AryTypePara[93].bit.sp := 16#0000;
   AryTypePara[93].bit.Other.Bool_1 := FALSE;
   AryTypePara[93].bit.Other.Byte_2 := 16#00;
   AryTypePara[93].bit.Other.Int_1 := 0;
   AryTypePara[93].bit.Other."Char" := ' ';
   AryTypePara[93].Other.STxxxCCDProgNO := 0;
   AryTypePara[93].Other.FixtureEnable := FALSE;
   AryTypePara[93].Other.Byte_1 := 16#00;
   AryTypePara[93].Other.Int_1 := 0;
   AryTypePara[93].Other."Char" := ' ';
   AryTypePara[93].Other.Word_1 := 16#0000;
   AryTypePara[93].Other.DInt_1 := 0;
   AryTypePara[93].Other.DWord_1 := 16#0000_0000;
   AryTypePara[93].Other.Real_1 := 0.0;
   AryTypePara[93].Other.S5Time := T#0MS;
   AryTypePara[93].Other."String" := '';
   AryTypePara[94].TypeName := '';
   AryTypePara[94].bit.Bit0 := FALSE;
   AryTypePara[94].bit.sp := 16#0000;
   AryTypePara[94].bit.Other.Bool_1 := FALSE;
   AryTypePara[94].bit.Other.Byte_2 := 16#00;
   AryTypePara[94].bit.Other.Int_1 := 0;
   AryTypePara[94].bit.Other."Char" := ' ';
   AryTypePara[94].Other.STxxxCCDProgNO := 0;
   AryTypePara[94].Other.FixtureEnable := FALSE;
   AryTypePara[94].Other.Byte_1 := 16#00;
   AryTypePara[94].Other.Int_1 := 0;
   AryTypePara[94].Other."Char" := ' ';
   AryTypePara[94].Other.Word_1 := 16#0000;
   AryTypePara[94].Other.DInt_1 := 0;
   AryTypePara[94].Other.DWord_1 := 16#0000_0000;
   AryTypePara[94].Other.Real_1 := 0.0;
   AryTypePara[94].Other.S5Time := T#0MS;
   AryTypePara[94].Other."String" := '';
   AryTypePara[95].TypeName := '';
   AryTypePara[95].bit.Bit0 := FALSE;
   AryTypePara[95].bit.sp := 16#0000;
   AryTypePara[95].bit.Other.Bool_1 := FALSE;
   AryTypePara[95].bit.Other.Byte_2 := 16#00;
   AryTypePara[95].bit.Other.Int_1 := 0;
   AryTypePara[95].bit.Other."Char" := ' ';
   AryTypePara[95].Other.STxxxCCDProgNO := 0;
   AryTypePara[95].Other.FixtureEnable := FALSE;
   AryTypePara[95].Other.Byte_1 := 16#00;
   AryTypePara[95].Other.Int_1 := 0;
   AryTypePara[95].Other."Char" := ' ';
   AryTypePara[95].Other.Word_1 := 16#0000;
   AryTypePara[95].Other.DInt_1 := 0;
   AryTypePara[95].Other.DWord_1 := 16#0000_0000;
   AryTypePara[95].Other.Real_1 := 0.0;
   AryTypePara[95].Other.S5Time := T#0MS;
   AryTypePara[95].Other."String" := '';
   AryTypePara[96].TypeName := '';
   AryTypePara[96].bit.Bit0 := FALSE;
   AryTypePara[96].bit.sp := 16#0000;
   AryTypePara[96].bit.Other.Bool_1 := FALSE;
   AryTypePara[96].bit.Other.Byte_2 := 16#00;
   AryTypePara[96].bit.Other.Int_1 := 0;
   AryTypePara[96].bit.Other."Char" := ' ';
   AryTypePara[96].Other.STxxxCCDProgNO := 0;
   AryTypePara[96].Other.FixtureEnable := FALSE;
   AryTypePara[96].Other.Byte_1 := 16#00;
   AryTypePara[96].Other.Int_1 := 0;
   AryTypePara[96].Other."Char" := ' ';
   AryTypePara[96].Other.Word_1 := 16#0000;
   AryTypePara[96].Other.DInt_1 := 0;
   AryTypePara[96].Other.DWord_1 := 16#0000_0000;
   AryTypePara[96].Other.Real_1 := 0.0;
   AryTypePara[96].Other.S5Time := T#0MS;
   AryTypePara[96].Other."String" := '';
   AryTypePara[97].TypeName := '';
   AryTypePara[97].bit.Bit0 := FALSE;
   AryTypePara[97].bit.sp := 16#0000;
   AryTypePara[97].bit.Other.Bool_1 := FALSE;
   AryTypePara[97].bit.Other.Byte_2 := 16#00;
   AryTypePara[97].bit.Other.Int_1 := 0;
   AryTypePara[97].bit.Other."Char" := ' ';
   AryTypePara[97].Other.STxxxCCDProgNO := 0;
   AryTypePara[97].Other.FixtureEnable := FALSE;
   AryTypePara[97].Other.Byte_1 := 16#00;
   AryTypePara[97].Other.Int_1 := 0;
   AryTypePara[97].Other."Char" := ' ';
   AryTypePara[97].Other.Word_1 := 16#0000;
   AryTypePara[97].Other.DInt_1 := 0;
   AryTypePara[97].Other.DWord_1 := 16#0000_0000;
   AryTypePara[97].Other.Real_1 := 0.0;
   AryTypePara[97].Other.S5Time := T#0MS;
   AryTypePara[97].Other."String" := '';
   AryTypePara[98].TypeName := '';
   AryTypePara[98].bit.Bit0 := FALSE;
   AryTypePara[98].bit.sp := 16#0000;
   AryTypePara[98].bit.Other.Bool_1 := FALSE;
   AryTypePara[98].bit.Other.Byte_2 := 16#00;
   AryTypePara[98].bit.Other.Int_1 := 0;
   AryTypePara[98].bit.Other."Char" := ' ';
   AryTypePara[98].Other.STxxxCCDProgNO := 0;
   AryTypePara[98].Other.FixtureEnable := FALSE;
   AryTypePara[98].Other.Byte_1 := 16#00;
   AryTypePara[98].Other.Int_1 := 0;
   AryTypePara[98].Other."Char" := ' ';
   AryTypePara[98].Other.Word_1 := 16#0000;
   AryTypePara[98].Other.DInt_1 := 0;
   AryTypePara[98].Other.DWord_1 := 16#0000_0000;
   AryTypePara[98].Other.Real_1 := 0.0;
   AryTypePara[98].Other.S5Time := T#0MS;
   AryTypePara[98].Other."String" := '';
   AryTypePara[99].TypeName := '';
   AryTypePara[99].bit.Bit0 := FALSE;
   AryTypePara[99].bit.sp := 16#0000;
   AryTypePara[99].bit.Other.Bool_1 := FALSE;
   AryTypePara[99].bit.Other.Byte_2 := 16#00;
   AryTypePara[99].bit.Other.Int_1 := 0;
   AryTypePara[99].bit.Other."Char" := ' ';
   AryTypePara[99].Other.STxxxCCDProgNO := 0;
   AryTypePara[99].Other.FixtureEnable := FALSE;
   AryTypePara[99].Other.Byte_1 := 16#00;
   AryTypePara[99].Other.Int_1 := 0;
   AryTypePara[99].Other."Char" := ' ';
   AryTypePara[99].Other.Word_1 := 16#0000;
   AryTypePara[99].Other.DInt_1 := 0;
   AryTypePara[99].Other.DWord_1 := 16#0000_0000;
   AryTypePara[99].Other.Real_1 := 0.0;
   AryTypePara[99].Other.S5Time := T#0MS;
   AryTypePara[99].Other."String" := '';
   AryTypePara[100].bit.Bit0 := FALSE;
   AryTypePara[100].bit.sp := 16#0000;
   AryTypePara[100].bit.Other.Bool_1 := FALSE;
   AryTypePara[100].bit.Other.Byte_2 := 16#00;
   AryTypePara[100].bit.Other.Int_1 := 0;
   AryTypePara[100].bit.Other."Char" := ' ';
   AryTypePara[100].Other.FixtureEnable := FALSE;
   AryTypePara[100].Other.Byte_1 := 16#00;
   AryTypePara[100].Other.Int_1 := 0;
   AryTypePara[100].Other."Char" := ' ';
   AryTypePara[100].Other.Word_1 := 16#0000;
   AryTypePara[100].Other.DInt_1 := 0;
   AryTypePara[100].Other.DWord_1 := 16#0000_0000;
   AryTypePara[100].Other.Real_1 := 0.0;
   AryTypePara[100].Other.S5Time := T#0MS;
   AryTypePara[100].Other."String" := '';
   AryTypePara[101].bit.Bit0 := FALSE;
   AryTypePara[101].bit.sp := 16#0000;
   AryTypePara[101].bit.Other.Bool_1 := FALSE;
   AryTypePara[101].bit.Other.Byte_2 := 16#00;
   AryTypePara[101].bit.Other.Int_1 := 0;
   AryTypePara[101].bit.Other."Char" := ' ';
   AryTypePara[101].Other.FixtureEnable := FALSE;
   AryTypePara[101].Other.Byte_1 := 16#00;
   AryTypePara[101].Other.Int_1 := 0;
   AryTypePara[101].Other."Char" := ' ';
   AryTypePara[101].Other.Word_1 := 16#0000;
   AryTypePara[101].Other.DInt_1 := 0;
   AryTypePara[101].Other.DWord_1 := 16#0000_0000;
   AryTypePara[101].Other.Real_1 := 0.0;
   AryTypePara[101].Other.S5Time := T#0MS;
   AryTypePara[101].Other."String" := '';
   AryTypePara[102].bit.Bit0 := FALSE;
   AryTypePara[102].bit.sp := 16#0000;
   AryTypePara[102].bit.Other.Bool_1 := FALSE;
   AryTypePara[102].bit.Other.Byte_2 := 16#00;
   AryTypePara[102].bit.Other.Int_1 := 0;
   AryTypePara[102].bit.Other."Char" := ' ';
   AryTypePara[102].Other.FixtureEnable := FALSE;
   AryTypePara[102].Other.Byte_1 := 16#00;
   AryTypePara[102].Other.Int_1 := 0;
   AryTypePara[102].Other."Char" := ' ';
   AryTypePara[102].Other.Word_1 := 16#0000;
   AryTypePara[102].Other.DInt_1 := 0;
   AryTypePara[102].Other.DWord_1 := 16#0000_0000;
   AryTypePara[102].Other.Real_1 := 0.0;
   AryTypePara[102].Other.S5Time := T#0MS;
   AryTypePara[102].Other."String" := '';
   AryTypePara[103].bit.Bit0 := FALSE;
   AryTypePara[103].bit.sp := 16#0000;
   AryTypePara[103].bit.Other.Bool_1 := FALSE;
   AryTypePara[103].bit.Other.Byte_2 := 16#00;
   AryTypePara[103].bit.Other.Int_1 := 0;
   AryTypePara[103].bit.Other."Char" := ' ';
   AryTypePara[103].Other.FixtureEnable := FALSE;
   AryTypePara[103].Other.Byte_1 := 16#00;
   AryTypePara[103].Other.Int_1 := 0;
   AryTypePara[103].Other."Char" := ' ';
   AryTypePara[103].Other.Word_1 := 16#0000;
   AryTypePara[103].Other.DInt_1 := 0;
   AryTypePara[103].Other.DWord_1 := 16#0000_0000;
   AryTypePara[103].Other.Real_1 := 0.0;
   AryTypePara[103].Other.S5Time := T#0MS;
   AryTypePara[103].Other."String" := '';
   AryTypePara[104].TypeName := '';
   AryTypePara[104].bit.Bit0 := FALSE;
   AryTypePara[104].bit.sp := 16#0000;
   AryTypePara[104].bit.Other.Bool_1 := FALSE;
   AryTypePara[104].bit.Other.Byte_2 := 16#00;
   AryTypePara[104].bit.Other.Int_1 := 0;
   AryTypePara[104].bit.Other."Char" := ' ';
   AryTypePara[104].Other.STxxxCCDProgNO := 0;
   AryTypePara[104].Other.FixtureEnable := FALSE;
   AryTypePara[104].Other.Byte_1 := 16#00;
   AryTypePara[104].Other.Int_1 := 0;
   AryTypePara[104].Other."Char" := ' ';
   AryTypePara[104].Other.Word_1 := 16#0000;
   AryTypePara[104].Other.DInt_1 := 0;
   AryTypePara[104].Other.DWord_1 := 16#0000_0000;
   AryTypePara[104].Other.Real_1 := 0.0;
   AryTypePara[104].Other.S5Time := T#0MS;
   AryTypePara[104].Other."String" := '';
   AryTypePara[105].TypeName := '';
   AryTypePara[105].bit.Bit0 := FALSE;
   AryTypePara[105].bit.sp := 16#0000;
   AryTypePara[105].bit.Other.Bool_1 := FALSE;
   AryTypePara[105].bit.Other.Byte_2 := 16#00;
   AryTypePara[105].bit.Other.Int_1 := 0;
   AryTypePara[105].bit.Other."Char" := ' ';
   AryTypePara[105].Other.STxxxCCDProgNO := 0;
